(* IEC 61131-3 sources: 2026_Projet_YGO_ExcavatriceDragage/TOOLS/TEST_AUTO_CI/RESULTS/L_SIMULATION/tests (part 7) *)

TEST 'TC-T418-INT-002 Refus puis retour permis sans nouvel appui'
nx := 5000; ny := 5000; raw1 := 0; raw2 := 0; previousButton := FALSE; buttonEdges := 0;
bench.Enable := TRUE; joy.Enable := TRUE; joy.ArmingPermit := TRUE; diagOk.Operational := TRUE;
joy.BusCanOpenOP := diagOk; joy.JoystickOP := diagOk; home.Enable := TRUE; home.BootReady := TRUE;
home.Mode := E_Mode.MAINT_N1; home.BucketOffsetValid := TRUE; home.WinchesMechanicallyStopped := TRUE;
joy.ArmingPermit := FALSE;
ADVANCE_TIME(10000000);
bench(RawPosM1 := raw1, RawPosM2 := raw2);
joy(RawX := bench.Operator.JoyXRaw_ANA1, RawY := bench.Operator.JoyYRaw_ANA2, RawButton := bench.Operator.JoyBtnRaw, Cfg := cfg, NeutralXMem := nx, NeutralYMem := ny);
home(DeadmanArmed := joy.DeadmanArmed, JoystickDeflected := NOT joy.AtNeutralXY, JoystickPull := joy.AxisCmdY.DirectionPositive, JoystickPush := joy.AxisCmdY.DirectionNegative, BtnValidation := bench.Operator.JoyBtnRaw);
IF bench.Operator.JoyBtnRaw AND NOT previousButton THEN buttonEdges := buttonEdges + 1; END_IF; previousButton := bench.Operator.JoyBtnRaw;
bench.SimJoystickFwd_Up_Close_Active := TRUE;
ADVANCE_TIME(10000000);
bench(RawPosM1 := raw1, RawPosM2 := raw2);
joy(RawX := bench.Operator.JoyXRaw_ANA1, RawY := bench.Operator.JoyYRaw_ANA2, RawButton := bench.Operator.JoyBtnRaw, Cfg := cfg, NeutralXMem := nx, NeutralYMem := ny);
home(DeadmanArmed := joy.DeadmanArmed, JoystickDeflected := NOT joy.AtNeutralXY, JoystickPull := joy.AxisCmdY.DirectionPositive, JoystickPush := joy.AxisCmdY.DirectionNegative, BtnValidation := bench.Operator.JoyBtnRaw);
IF bench.Operator.JoyBtnRaw AND NOT previousButton THEN buttonEdges := buttonEdges + 1; END_IF; previousButton := bench.Operator.JoyBtnRaw;
ASSERT_FALSE(joy.AxisCmdY.StartStop, 'Permis absent aucun mouvement'); ASSERT_FALSE(joy.DeadmanArmed, 'Refus reel');
ADVANCE_TIME(10000000);
bench(RawPosM1 := raw1, RawPosM2 := raw2);
joy(RawX := bench.Operator.JoyXRaw_ANA1, RawY := bench.Operator.JoyYRaw_ANA2, RawButton := bench.Operator.JoyBtnRaw, Cfg := cfg, NeutralXMem := nx, NeutralYMem := ny);
home(DeadmanArmed := joy.DeadmanArmed, JoystickDeflected := NOT joy.AtNeutralXY, JoystickPull := joy.AxisCmdY.DirectionPositive, JoystickPush := joy.AxisCmdY.DirectionNegative, BtnValidation := bench.Operator.JoyBtnRaw);
IF bench.Operator.JoyBtnRaw AND NOT previousButton THEN buttonEdges := buttonEdges + 1; END_IF; previousButton := bench.Operator.JoyBtnRaw;
ASSERT_FALSE(joy.AxisCmdY.StartStop, 'Permis absent aucun mouvement'); ASSERT_FALSE(joy.DeadmanArmed, 'Refus reel');
ADVANCE_TIME(10000000);
bench(RawPosM1 := raw1, RawPosM2 := raw2);
joy(RawX := bench.Operator.JoyXRaw_ANA1, RawY := bench.Operator.JoyYRaw_ANA2, RawButton := bench.Operator.JoyBtnRaw, Cfg := cfg, NeutralXMem := nx, NeutralYMem := ny);
home(DeadmanArmed := joy.DeadmanArmed, JoystickDeflected := NOT joy.AtNeutralXY, JoystickPull := joy.AxisCmdY.DirectionPositive, JoystickPush := joy.AxisCmdY.DirectionNegative, BtnValidation := bench.Operator.JoyBtnRaw);
IF bench.Operator.JoyBtnRaw AND NOT previousButton THEN buttonEdges := buttonEdges + 1; END_IF; previousButton := bench.Operator.JoyBtnRaw;
ASSERT_FALSE(joy.AxisCmdY.StartStop, 'Permis absent aucun mouvement'); ASSERT_FALSE(joy.DeadmanArmed, 'Refus reel');
ADVANCE_TIME(10000000);
bench(RawPosM1 := raw1, RawPosM2 := raw2);
joy(RawX := bench.Operator.JoyXRaw_ANA1, RawY := bench.Operator.JoyYRaw_ANA2, RawButton := bench.Operator.JoyBtnRaw, Cfg := cfg, NeutralXMem := nx, NeutralYMem := ny);
home(DeadmanArmed := joy.DeadmanArmed, JoystickDeflected := NOT joy.AtNeutralXY, JoystickPull := joy.AxisCmdY.DirectionPositive, JoystickPush := joy.AxisCmdY.DirectionNegative, BtnValidation := bench.Operator.JoyBtnRaw);
IF bench.Operator.JoyBtnRaw AND NOT previousButton THEN buttonEdges := buttonEdges + 1; END_IF; previousButton := bench.Operator.JoyBtnRaw;
ASSERT_FALSE(joy.AxisCmdY.StartStop, 'Permis absent aucun mouvement'); ASSERT_FALSE(joy.DeadmanArmed, 'Refus reel');
ADVANCE_TIME(10000000);
bench(RawPosM1 := raw1, RawPosM2 := raw2);
joy(RawX := bench.Operator.JoyXRaw_ANA1, RawY := bench.Operator.JoyYRaw_ANA2, RawButton := bench.Operator.JoyBtnRaw, Cfg := cfg, NeutralXMem := nx, NeutralYMem := ny);
home(DeadmanArmed := joy.DeadmanArmed, JoystickDeflected := NOT joy.AtNeutralXY, JoystickPull := joy.AxisCmdY.DirectionPositive, JoystickPush := joy.AxisCmdY.DirectionNegative, BtnValidation := bench.Operator.JoyBtnRaw);
IF bench.Operator.JoyBtnRaw AND NOT previousButton THEN buttonEdges := buttonEdges + 1; END_IF; previousButton := bench.Operator.JoyBtnRaw;
ASSERT_FALSE(joy.AxisCmdY.StartStop, 'Permis absent aucun mouvement'); ASSERT_FALSE(joy.DeadmanArmed, 'Refus reel');
ADVANCE_TIME(10000000);
bench(RawPosM1 := raw1, RawPosM2 := raw2);
joy(RawX := bench.Operator.JoyXRaw_ANA1, RawY := bench.Operator.JoyYRaw_ANA2, RawButton := bench.Operator.JoyBtnRaw, Cfg := cfg, NeutralXMem := nx, NeutralYMem := ny);
home(DeadmanArmed := joy.DeadmanArmed, JoystickDeflected := NOT joy.AtNeutralXY, JoystickPull := joy.AxisCmdY.DirectionPositive, JoystickPush := joy.AxisCmdY.DirectionNegative, BtnValidation := bench.Operator.JoyBtnRaw);
IF bench.Operator.JoyBtnRaw AND NOT previousButton THEN buttonEdges := buttonEdges + 1; END_IF; previousButton := bench.Operator.JoyBtnRaw;
ASSERT_FALSE(joy.AxisCmdY.StartStop, 'Permis absent aucun mouvement'); ASSERT_FALSE(joy.DeadmanArmed, 'Refus reel');
ADVANCE_TIME(10000000);
bench(RawPosM1 := raw1, RawPosM2 := raw2);
joy(RawX := bench.Operator.JoyXRaw_ANA1, RawY := bench.Operator.JoyYRaw_ANA2, RawButton := bench.Operator.JoyBtnRaw, Cfg := cfg, NeutralXMem := nx, NeutralYMem := ny);
home(DeadmanArmed := joy.DeadmanArmed, JoystickDeflected := NOT joy.AtNeutralXY, JoystickPull := joy.AxisCmdY.DirectionPositive, JoystickPush := joy.AxisCmdY.DirectionNegative, BtnValidation := bench.Operator.JoyBtnRaw);
IF bench.Operator.JoyBtnRaw AND NOT previousButton THEN buttonEdges := buttonEdges + 1; END_IF; previousButton := bench.Operator.JoyBtnRaw;
ASSERT_FALSE(joy.AxisCmdY.StartStop, 'Permis absent aucun mouvement'); ASSERT_FALSE(joy.DeadmanArmed, 'Refus reel');
ADVANCE_TIME(10000000);
bench(RawPosM1 := raw1, RawPosM2 := raw2);
joy(RawX := bench.Operator.JoyXRaw_ANA1, RawY := bench.Operator.JoyYRaw_ANA2, RawButton := bench.Operator.JoyBtnRaw, Cfg := cfg, NeutralXMem := nx, NeutralYMem := ny);
home(DeadmanArmed := joy.DeadmanArmed, JoystickDeflected := NOT joy.AtNeutralXY, JoystickPull := joy.AxisCmdY.DirectionPositive, JoystickPush := joy.AxisCmdY.DirectionNegative, BtnValidation := bench.Operator.JoyBtnRaw);
IF bench.Operator.JoyBtnRaw AND NOT previousButton THEN buttonEdges := buttonEdges + 1; END_IF; previousButton := bench.Operator.JoyBtnRaw;
ASSERT_FALSE(joy.AxisCmdY.StartStop, 'Permis absent aucun mouvement'); ASSERT_FALSE(joy.DeadmanArmed, 'Refus reel');
ADVANCE_TIME(10000000);
bench(RawPosM1 := raw1, RawPosM2 := raw2);
joy(RawX := bench.Operator.JoyXRaw_ANA1, RawY := bench.Operator.JoyYRaw_ANA2, RawButton := bench.Operator.JoyBtnRaw, Cfg := cfg, NeutralXMem := nx, NeutralYMem := ny);
home(DeadmanArmed := joy.DeadmanArmed, JoystickDeflected := NOT joy.AtNeutralXY, JoystickPull := joy.AxisCmdY.DirectionPositive, JoystickPush := joy.AxisCmdY.DirectionNegative, BtnValidation := bench.Operator.JoyBtnRaw);
IF bench.Operator.JoyBtnRaw AND NOT previousButton THEN buttonEdges := buttonEdges + 1; END_IF; previousButton := bench.Operator.JoyBtnRaw;
ASSERT_FALSE(joy.AxisCmdY.StartStop, 'Permis absent aucun mouvement'); ASSERT_FALSE(joy.DeadmanArmed, 'Refus reel');
ADVANCE_TIME(10000000);
bench(RawPosM1 := raw1, RawPosM2 := raw2);
joy(RawX := bench.Operator.JoyXRaw_ANA1, RawY := bench.Operator.JoyYRaw_ANA2, RawButton := bench.Operator.JoyBtnRaw, Cfg := cfg, NeutralXMem := nx, NeutralYMem := ny);
home(DeadmanArmed := joy.DeadmanArmed, JoystickDeflected := NOT joy.AtNeutralXY, JoystickPull := joy.AxisCmdY.DirectionPositive, JoystickPush := joy.AxisCmdY.DirectionNegative, BtnValidation := bench.Operator.JoyBtnRaw);
IF bench.Operator.JoyBtnRaw AND NOT previousButton THEN buttonEdges := buttonEdges + 1; END_IF; previousButton := bench.Operator.JoyBtnRaw;
ASSERT_FALSE(joy.AxisCmdY.StartStop, 'Permis absent aucun mouvement'); ASSERT_FALSE(joy.DeadmanArmed, 'Refus reel');
ADVANCE_TIME(10000000);
bench(RawPosM1 := raw1, RawPosM2 := raw2);
joy(RawX := bench.Operator.JoyXRaw_ANA1, RawY := bench.Operator.JoyYRaw_ANA2, RawButton := bench.Operator.JoyBtnRaw, Cfg := cfg, NeutralXMem := nx, NeutralYMem := ny);
home(DeadmanArmed := joy.DeadmanArmed, JoystickDeflected := NOT joy.AtNeutralXY, JoystickPull := joy.AxisCmdY.DirectionPositive, JoystickPush := joy.AxisCmdY.DirectionNegative, BtnValidation := bench.Operator.JoyBtnRaw);
IF bench.Operator.JoyBtnRaw AND NOT previousButton THEN buttonEdges := buttonEdges + 1; END_IF; previousButton := bench.Operator.JoyBtnRaw;
ASSERT_FALSE(joy.AxisCmdY.StartStop, 'Permis absent aucun mouvement'); ASSERT_FALSE(joy.DeadmanArmed, 'Refus reel');
ADVANCE_TIME(10000000);
bench(RawPosM1 := raw1, RawPosM2 := raw2);
joy(RawX := bench.Operator.JoyXRaw_ANA1, RawY := bench.Operator.JoyYRaw_ANA2, RawButton := bench.Operator.JoyBtnRaw, Cfg := cfg, NeutralXMem := nx, NeutralYMem := ny);
home(DeadmanArmed := joy.DeadmanArmed, JoystickDeflected := NOT joy.AtNeutralXY, JoystickPull := joy.AxisCmdY.DirectionPositive, JoystickPush := joy.AxisCmdY.DirectionNegative, BtnValidation := bench.Operator.JoyBtnRaw);
IF bench.Operator.JoyBtnRaw AND NOT previousButton THEN buttonEdges := buttonEdges + 1; END_IF; previousButton := bench.Operator.JoyBtnRaw;
ASSERT_FALSE(joy.AxisCmdY.StartStop, 'Permis absent aucun mouvement'); ASSERT_FALSE(joy.DeadmanArmed, 'Refus reel');
ADVANCE_TIME(10000000);
bench(RawPosM1 := raw1, RawPosM2 := raw2);
joy(RawX := bench.Operator.JoyXRaw_ANA1, RawY := bench.Operator.JoyYRaw_ANA2, RawButton := bench.Operator.JoyBtnRaw, Cfg := cfg, NeutralXMem := nx, NeutralYMem := ny);
home(DeadmanArmed := joy.DeadmanArmed, JoystickDeflected := NOT joy.AtNeutralXY, JoystickPull := joy.AxisCmdY.DirectionPositive, JoystickPush := joy.AxisCmdY.DirectionNegative, BtnValidation := bench.Operator.JoyBtnRaw);
IF bench.Operator.JoyBtnRaw AND NOT previousButton THEN buttonEdges := buttonEdges + 1; END_IF; previousButton := bench.Operator.JoyBtnRaw;
ASSERT_FALSE(joy.AxisCmdY.StartStop, 'Permis absent aucun mouvement'); ASSERT_FALSE(joy.DeadmanArmed, 'Refus reel');
ADVANCE_TIME(10000000);
bench(RawPosM1 := raw1, RawPosM2 := raw2);
joy(RawX := bench.Operator.JoyXRaw_ANA1, RawY := bench.Operator.JoyYRaw_ANA2, RawButton := bench.Operator.JoyBtnRaw, Cfg := cfg, NeutralXMem := nx, NeutralYMem := ny);
home(DeadmanArmed := joy.DeadmanArmed, JoystickDeflected := NOT joy.AtNeutralXY, JoystickPull := joy.AxisCmdY.DirectionPositive, JoystickPush := joy.AxisCmdY.DirectionNegative, BtnValidation := bench.Operator.JoyBtnRaw);
IF bench.Operator.JoyBtnRaw AND NOT previousButton THEN buttonEdges := buttonEdges + 1; END_IF; previousButton := bench.Operator.JoyBtnRaw;
ASSERT_FALSE(joy.AxisCmdY.StartStop, 'Permis absent aucun mouvement'); ASSERT_FALSE(joy.DeadmanArmed, 'Refus reel');
ADVANCE_TIME(10000000);
bench(RawPosM1 := raw1, RawPosM2 := raw2);
joy(RawX := bench.Operator.JoyXRaw_ANA1, RawY := bench.Operator.JoyYRaw_ANA2, RawButton := bench.Operator.JoyBtnRaw, Cfg := cfg, NeutralXMem := nx, NeutralYMem := ny);
home(DeadmanArmed := joy.DeadmanArmed, JoystickDeflected := NOT joy.AtNeutralXY, JoystickPull := joy.AxisCmdY.DirectionPositive, JoystickPush := joy.AxisCmdY.DirectionNegative, BtnValidation := bench.Operator.JoyBtnRaw);
IF bench.Operator.JoyBtnRaw AND NOT previousButton THEN buttonEdges := buttonEdges + 1; END_IF; previousButton := bench.Operator.JoyBtnRaw;
ASSERT_FALSE(joy.AxisCmdY.StartStop, 'Permis absent aucun mouvement'); ASSERT_FALSE(joy.DeadmanArmed, 'Refus reel');
ADVANCE_TIME(10000000);
bench(RawPosM1 := raw1, RawPosM2 := raw2);
joy(RawX := bench.Operator.JoyXRaw_ANA1, RawY := bench.Operator.JoyYRaw_ANA2, RawButton := bench.Operator.JoyBtnRaw, Cfg := cfg, NeutralXMem := nx, NeutralYMem := ny);
home(DeadmanArmed := joy.DeadmanArmed, JoystickDeflected := NOT joy.AtNeutralXY, JoystickPull := joy.AxisCmdY.DirectionPositive, JoystickPush := joy.AxisCmdY.DirectionNegative, BtnValidation := bench.Operator.JoyBtnRaw);
IF bench.Operator.JoyBtnRaw AND NOT previousButton THEN buttonEdges := buttonEdges + 1; END_IF; previousButton := bench.Operator.JoyBtnRaw;
ASSERT_FALSE(joy.AxisCmdY.StartStop, 'Permis absent aucun mouvement'); ASSERT_FALSE(joy.DeadmanArmed, 'Refus reel');
ADVANCE_TIME(10000000);
bench(RawPosM1 := raw1, RawPosM2 := raw2);
joy(RawX := bench.Operator.JoyXRaw_ANA1, RawY := bench.Operator.JoyYRaw_ANA2, RawButton := bench.Operator.JoyBtnRaw, Cfg := cfg, NeutralXMem := nx, NeutralYMem := ny);
home(DeadmanArmed := joy.DeadmanArmed, JoystickDeflected := NOT joy.AtNeutralXY, JoystickPull := joy.AxisCmdY.DirectionPositive, JoystickPush := joy.AxisCmdY.DirectionNegative, BtnValidation := bench.Operator.JoyBtnRaw);
IF bench.Operator.JoyBtnRaw AND NOT previousButton THEN buttonEdges := buttonEdges + 1; END_IF; previousButton := bench.Operator.JoyBtnRaw;
ASSERT_FALSE(joy.AxisCmdY.StartStop, 'Permis absent aucun mouvement'); ASSERT_FALSE(joy.DeadmanArmed, 'Refus reel');
ADVANCE_TIME(10000000);
bench(RawPosM1 := raw1, RawPosM2 := raw2);
joy(RawX := bench.Operator.JoyXRaw_ANA1, RawY := bench.Operator.JoyYRaw_ANA2, RawButton := bench.Operator.JoyBtnRaw, Cfg := cfg, NeutralXMem := nx, NeutralYMem := ny);
home(DeadmanArmed := joy.DeadmanArmed, JoystickDeflected := NOT joy.AtNeutralXY, JoystickPull := joy.AxisCmdY.DirectionPositive, JoystickPush := joy.AxisCmdY.DirectionNegative, BtnValidation := bench.Operator.JoyBtnRaw);
IF bench.Operator.JoyBtnRaw AND NOT previousButton THEN buttonEdges := buttonEdges + 1; END_IF; previousButton := bench.Operator.JoyBtnRaw;
ASSERT_FALSE(joy.AxisCmdY.StartStop, 'Permis absent aucun mouvement'); ASSERT_FALSE(joy.DeadmanArmed, 'Refus reel');
ADVANCE_TIME(10000000);
bench(RawPosM1 := raw1, RawPosM2 := raw2);
joy(RawX := bench.Operator.JoyXRaw_ANA1, RawY := bench.Operator.JoyYRaw_ANA2, RawButton := bench.Operator.JoyBtnRaw, Cfg := cfg, NeutralXMem := nx, NeutralYMem := ny);
home(DeadmanArmed := joy.DeadmanArmed, JoystickDeflected := NOT joy.AtNeutralXY, JoystickPull := joy.AxisCmdY.DirectionPositive, JoystickPush := joy.AxisCmdY.DirectionNegative, BtnValidation := bench.Operator.JoyBtnRaw);
IF bench.Operator.JoyBtnRaw AND NOT previousButton THEN buttonEdges := buttonEdges + 1; END_IF; previousButton := bench.Operator.JoyBtnRaw;
ASSERT_FALSE(joy.AxisCmdY.StartStop, 'Permis absent aucun mouvement'); ASSERT_FALSE(joy.DeadmanArmed, 'Refus reel');
ADVANCE_TIME(10000000);
bench(RawPosM1 := raw1, RawPosM2 := raw2);
joy(RawX := bench.Operator.JoyXRaw_ANA1, RawY := bench.Operator.JoyYRaw_ANA2, RawButton := bench.Operator.JoyBtnRaw, Cfg := cfg, NeutralXMem := nx, NeutralYMem := ny);
home(DeadmanArmed := joy.DeadmanArmed, JoystickDeflected := NOT joy.AtNeutralXY, JoystickPull := joy.AxisCmdY.DirectionPositive, JoystickPush := joy.AxisCmdY.DirectionNegative, BtnValidation := bench.Operator.JoyBtnRaw);
IF bench.Operator.JoyBtnRaw AND NOT previousButton THEN buttonEdges := buttonEdges + 1; END_IF; previousButton := bench.Operator.JoyBtnRaw;
ASSERT_FALSE(joy.AxisCmdY.StartStop, 'Permis absent aucun mouvement'); ASSERT_FALSE(joy.DeadmanArmed, 'Refus reel');
ADVANCE_TIME(10000000);
bench(RawPosM1 := raw1, RawPosM2 := raw2);
joy(RawX := bench.Operator.JoyXRaw_ANA1, RawY := bench.Operator.JoyYRaw_ANA2, RawButton := bench.Operator.JoyBtnRaw, Cfg := cfg, NeutralXMem := nx, NeutralYMem := ny);
home(DeadmanArmed := joy.DeadmanArmed, JoystickDeflected := NOT joy.AtNeutralXY, JoystickPull := joy.AxisCmdY.DirectionPositive, JoystickPush := joy.AxisCmdY.DirectionNegative, BtnValidation := bench.Operator.JoyBtnRaw);
IF bench.Operator.JoyBtnRaw AND NOT previousButton THEN buttonEdges := buttonEdges + 1; END_IF; previousButton := bench.Operator.JoyBtnRaw;
ASSERT_FALSE(joy.AxisCmdY.StartStop, 'Permis absent aucun mouvement'); ASSERT_FALSE(joy.DeadmanArmed, 'Refus reel');
ADVANCE_TIME(10000000);
bench(RawPosM1 := raw1, RawPosM2 := raw2);
joy(RawX := bench.Operator.JoyXRaw_ANA1, RawY := bench.Operator.JoyYRaw_ANA2, RawButton := bench.Operator.JoyBtnRaw, Cfg := cfg, NeutralXMem := nx, NeutralYMem := ny);
home(DeadmanArmed := joy.DeadmanArmed, JoystickDeflected := NOT joy.AtNeutralXY, JoystickPull := joy.AxisCmdY.DirectionPositive, JoystickPush := joy.AxisCmdY.DirectionNegative, BtnValidation := bench.Operator.JoyBtnRaw);
IF bench.Operator.JoyBtnRaw AND NOT previousButton THEN buttonEdges := buttonEdges + 1; END_IF; previousButton := bench.Operator.JoyBtnRaw;
ASSERT_FALSE(joy.AxisCmdY.StartStop, 'Permis absent aucun mouvement'); ASSERT_FALSE(joy.DeadmanArmed, 'Refus reel');
ADVANCE_TIME(10000000);
bench(RawPosM1 := raw1, RawPosM2 := raw2);
joy(RawX := bench.Operator.JoyXRaw_ANA1, RawY := bench.Operator.JoyYRaw_ANA2, RawButton := bench.Operator.JoyBtnRaw, Cfg := cfg, NeutralXMem := nx, NeutralYMem := ny);
home(DeadmanArmed := joy.DeadmanArmed, JoystickDeflected := NOT joy.AtNeutralXY, JoystickPull := joy.AxisCmdY.DirectionPositive, JoystickPush := joy.AxisCmdY.DirectionNegative, BtnValidation := bench.Operator.JoyBtnRaw);
IF bench.Operator.JoyBtnRaw AND NOT previousButton THEN buttonEdges := buttonEdges + 1; END_IF; previousButton := bench.Operator.JoyBtnRaw;
ASSERT_FALSE(joy.AxisCmdY.StartStop, 'Permis absent aucun mouvement'); ASSERT_FALSE(joy.DeadmanArmed, 'Refus reel');
ADVANCE_TIME(10000000);
bench(RawPosM1 := raw1, RawPosM2 := raw2);
joy(RawX := bench.Operator.JoyXRaw_ANA1, RawY := bench.Operator.JoyYRaw_ANA2, RawButton := bench.Operator.JoyBtnRaw, Cfg := cfg, NeutralXMem := nx, NeutralYMem := ny);
home(DeadmanArmed := joy.DeadmanArmed, JoystickDeflected := NOT joy.AtNeutralXY, JoystickPull := joy.AxisCmdY.DirectionPositive, JoystickPush := joy.AxisCmdY.DirectionNegative, BtnValidation := bench.Operator.JoyBtnRaw);
IF bench.Operator.JoyBtnRaw AND NOT previousButton THEN buttonEdges := buttonEdges + 1; END_IF; previousButton := bench.Operator.JoyBtnRaw;
ASSERT_FALSE(joy.AxisCmdY.StartStop, 'Permis absent aucun mouvement'); ASSERT_FALSE(joy.DeadmanArmed, 'Refus reel');
ADVANCE_TIME(10000000);
bench(RawPosM1 := raw1, RawPosM2 := raw2);
joy(RawX := bench.Operator.JoyXRaw_ANA1, RawY := bench.Operator.JoyYRaw_ANA2, RawButton := bench.Operator.JoyBtnRaw, Cfg := cfg, NeutralXMem := nx, NeutralYMem := ny);
home(DeadmanArmed := joy.DeadmanArmed, JoystickDeflected := NOT joy.AtNeutralXY, JoystickPull := joy.AxisCmdY.DirectionPositive, JoystickPush := joy.AxisCmdY.DirectionNegative, BtnValidation := bench.Operator.JoyBtnRaw);
IF bench.Operator.JoyBtnRaw AND NOT previousButton THEN buttonEdges := buttonEdges + 1; END_IF; previousButton := bench.Operator.JoyBtnRaw;
ASSERT_FALSE(joy.AxisCmdY.StartStop, 'Permis absent aucun mouvement'); ASSERT_FALSE(joy.DeadmanArmed, 'Refus reel');
ADVANCE_TIME(10000000);
bench(RawPosM1 := raw1, RawPosM2 := raw2);
joy(RawX := bench.Operator.JoyXRaw_ANA1, RawY := bench.Operator.JoyYRaw_ANA2, RawButton := bench.Operator.JoyBtnRaw, Cfg := cfg, NeutralXMem := nx, NeutralYMem := ny);
home(DeadmanArmed := joy.DeadmanArmed, JoystickDeflected := NOT joy.AtNeutralXY, JoystickPull := joy.AxisCmdY.DirectionPositive, JoystickPush := joy.AxisCmdY.DirectionNegative, BtnValidation := bench.Operator.JoyBtnRaw);
IF bench.Operator.JoyBtnRaw AND NOT previousButton THEN buttonEdges := buttonEdges + 1; END_IF; previousButton := bench.Operator.JoyBtnRaw;
ASSERT_FALSE(joy.AxisCmdY.StartStop, 'Permis absent aucun mouvement'); ASSERT_FALSE(joy.DeadmanArmed, 'Refus reel');
ADVANCE_TIME(10000000);
bench(RawPosM1 := raw1, RawPosM2 := raw2);
joy(RawX := bench.Operator.JoyXRaw_ANA1, RawY := bench.Operator.JoyYRaw_ANA2, RawButton := bench.Operator.JoyBtnRaw, Cfg := cfg, NeutralXMem := nx, NeutralYMem := ny);
home(DeadmanArmed := joy.DeadmanArmed, JoystickDeflected := NOT joy.AtNeutralXY, JoystickPull := joy.AxisCmdY.DirectionPositive, JoystickPush := joy.AxisCmdY.DirectionNegative, BtnValidation := bench.Operator.JoyBtnRaw);
IF bench.Operator.JoyBtnRaw AND NOT previousButton THEN buttonEdges := buttonEdges + 1; END_IF; previousButton := bench.Operator.JoyBtnRaw;
ASSERT_FALSE(joy.AxisCmdY.StartStop, 'Permis absent aucun mouvement'); ASSERT_FALSE(joy.DeadmanArmed, 'Refus reel');
ADVANCE_TIME(10000000);
bench(RawPosM1 := raw1, RawPosM2 := raw2);
joy(RawX := bench.Operator.JoyXRaw_ANA1, RawY := bench.Operator.JoyYRaw_ANA2, RawButton := bench.Operator.JoyBtnRaw, Cfg := cfg, NeutralXMem := nx, NeutralYMem := ny);
home(DeadmanArmed := joy.DeadmanArmed, JoystickDeflected := NOT joy.AtNeutralXY, JoystickPull := joy.AxisCmdY.DirectionPositive, JoystickPush := joy.AxisCmdY.DirectionNegative, BtnValidation := bench.Operator.JoyBtnRaw);
IF bench.Operator.JoyBtnRaw AND NOT previousButton THEN buttonEdges := buttonEdges + 1; END_IF; previousButton := bench.Operator.JoyBtnRaw;
ASSERT_FALSE(joy.AxisCmdY.StartStop, 'Permis absent aucun mouvement'); ASSERT_FALSE(joy.DeadmanArmed, 'Refus reel');
ADVANCE_TIME(10000000);
bench(RawPosM1 := raw1, RawPosM2 := raw2);
joy(RawX := bench.Operator.JoyXRaw_ANA1, RawY := bench.Operator.JoyYRaw_ANA2, RawButton := bench.Operator.JoyBtnRaw, Cfg := cfg, NeutralXMem := nx, NeutralYMem := ny);
home(DeadmanArmed := joy.DeadmanArmed, JoystickDeflected := NOT joy.AtNeutralXY, JoystickPull := joy.AxisCmdY.DirectionPositive, JoystickPush := joy.AxisCmdY.DirectionNegative, BtnValidation := bench.Operator.JoyBtnRaw);
IF bench.Operator.JoyBtnRaw AND NOT previousButton THEN buttonEdges := buttonEdges + 1; END_IF; previousButton := bench.Operator.JoyBtnRaw;
ASSERT_FALSE(joy.AxisCmdY.StartStop, 'Permis absent aucun mouvement'); ASSERT_FALSE(joy.DeadmanArmed, 'Refus reel');
ADVANCE_TIME(10000000);
bench(RawPosM1 := raw1, RawPosM2 := raw2);
joy(RawX := bench.Operator.JoyXRaw_ANA1, RawY := bench.Operator.JoyYRaw_ANA2, RawButton := bench.Operator.JoyBtnRaw, Cfg := cfg, NeutralXMem := nx, NeutralYMem := ny);
home(DeadmanArmed := joy.DeadmanArmed, JoystickDeflected := NOT joy.AtNeutralXY, JoystickPull := joy.AxisCmdY.DirectionPositive, JoystickPush := joy.AxisCmdY.DirectionNegative, BtnValidation := bench.Operator.JoyBtnRaw);
IF bench.Operator.JoyBtnRaw AND NOT previousButton THEN buttonEdges := buttonEdges + 1; END_IF; previousButton := bench.Operator.JoyBtnRaw;
ASSERT_FALSE(joy.AxisCmdY.StartStop, 'Permis absent aucun mouvement'); ASSERT_FALSE(joy.DeadmanArmed, 'Refus reel');
ADVANCE_TIME(10000000);
bench(RawPosM1 := raw1, RawPosM2 := raw2);
joy(RawX := bench.Operator.JoyXRaw_ANA1, RawY := bench.Operator.JoyYRaw_ANA2, RawButton := bench.Operator.JoyBtnRaw, Cfg := cfg, NeutralXMem := nx, NeutralYMem := ny);
home(DeadmanArmed := joy.DeadmanArmed, JoystickDeflected := NOT joy.AtNeutralXY, JoystickPull := joy.AxisCmdY.DirectionPositive, JoystickPush := joy.AxisCmdY.DirectionNegative, BtnValidation := bench.Operator.JoyBtnRaw);
IF bench.Operator.JoyBtnRaw AND NOT previousButton THEN buttonEdges := buttonEdges + 1; END_IF; previousButton := bench.Operator.JoyBtnRaw;
ASSERT_FALSE(joy.AxisCmdY.StartStop, 'Permis absent aucun mouvement'); ASSERT_FALSE(joy.DeadmanArmed, 'Refus reel');
ADVANCE_TIME(10000000);
bench(RawPosM1 := raw1, RawPosM2 := raw2);
joy(RawX := bench.Operator.JoyXRaw_ANA1, RawY := bench.Operator.JoyYRaw_ANA2, RawButton := bench.Operator.JoyBtnRaw, Cfg := cfg, NeutralXMem := nx, NeutralYMem := ny);
home(DeadmanArmed := joy.DeadmanArmed, JoystickDeflected := NOT joy.AtNeutralXY, JoystickPull := joy.AxisCmdY.DirectionPositive, JoystickPush := joy.AxisCmdY.DirectionNegative, BtnValidation := bench.Operator.JoyBtnRaw);
IF bench.Operator.JoyBtnRaw AND NOT previousButton THEN buttonEdges := buttonEdges + 1; END_IF; previousButton := bench.Operator.JoyBtnRaw;
ASSERT_FALSE(joy.AxisCmdY.StartStop, 'Permis absent aucun mouvement'); ASSERT_FALSE(joy.DeadmanArmed, 'Refus reel');
ADVANCE_TIME(10000000);
bench(RawPosM1 := raw1, RawPosM2 := raw2);
joy(RawX := bench.Operator.JoyXRaw_ANA1, RawY := bench.Operator.JoyYRaw_ANA2, RawButton := bench.Operator.JoyBtnRaw, Cfg := cfg, NeutralXMem := nx, NeutralYMem := ny);
home(DeadmanArmed := joy.DeadmanArmed, JoystickDeflected := NOT joy.AtNeutralXY, JoystickPull := joy.AxisCmdY.DirectionPositive, JoystickPush := joy.AxisCmdY.DirectionNegative, BtnValidation := bench.Operator.JoyBtnRaw);
IF bench.Operator.JoyBtnRaw AND NOT previousButton THEN buttonEdges := buttonEdges + 1; END_IF; previousButton := bench.Operator.JoyBtnRaw;
ASSERT_FALSE(joy.AxisCmdY.StartStop, 'Permis absent aucun mouvement'); ASSERT_FALSE(joy.DeadmanArmed, 'Refus reel');
ADVANCE_TIME(10000000);
bench(RawPosM1 := raw1, RawPosM2 := raw2);
joy(RawX := bench.Operator.JoyXRaw_ANA1, RawY := bench.Operator.JoyYRaw_ANA2, RawButton := bench.Operator.JoyBtnRaw, Cfg := cfg, NeutralXMem := nx, NeutralYMem := ny);
home(DeadmanArmed := joy.DeadmanArmed, JoystickDeflected := NOT joy.AtNeutralXY, JoystickPull := joy.AxisCmdY.DirectionPositive, JoystickPush := joy.AxisCmdY.DirectionNegative, BtnValidation := bench.Operator.JoyBtnRaw);
IF bench.Operator.JoyBtnRaw AND NOT previousButton THEN buttonEdges := buttonEdges + 1; END_IF; previousButton := bench.Operator.JoyBtnRaw;
ASSERT_FALSE(joy.AxisCmdY.StartStop, 'Permis absent aucun mouvement'); ASSERT_FALSE(joy.DeadmanArmed, 'Refus reel');
ADVANCE_TIME(10000000);
bench(RawPosM1 := raw1, RawPosM2 := raw2);
joy(RawX := bench.Operator.JoyXRaw_ANA1, RawY := bench.Operator.JoyYRaw_ANA2, RawButton := bench.Operator.JoyBtnRaw, Cfg := cfg, NeutralXMem := nx, NeutralYMem := ny);
home(DeadmanArmed := joy.DeadmanArmed, JoystickDeflected := NOT joy.AtNeutralXY, JoystickPull := joy.AxisCmdY.DirectionPositive, JoystickPush := joy.AxisCmdY.DirectionNegative, BtnValidation := bench.Operator.JoyBtnRaw);
IF bench.Operator.JoyBtnRaw AND NOT previousButton THEN buttonEdges := buttonEdges + 1; END_IF; previousButton := bench.Operator.JoyBtnRaw;
ASSERT_FALSE(joy.AxisCmdY.StartStop, 'Permis absent aucun mouvement'); ASSERT_FALSE(joy.DeadmanArmed, 'Refus reel');
ADVANCE_TIME(10000000);
bench(RawPosM1 := raw1, RawPosM2 := raw2);
joy(RawX := bench.Operator.JoyXRaw_ANA1, RawY := bench.Operator.JoyYRaw_ANA2, RawButton := bench.Operator.JoyBtnRaw, Cfg := cfg, NeutralXMem := nx, NeutralYMem := ny);
home(DeadmanArmed := joy.DeadmanArmed, JoystickDeflected := NOT joy.AtNeutralXY, JoystickPull := joy.AxisCmdY.DirectionPositive, JoystickPush := joy.AxisCmdY.DirectionNegative, BtnValidation := bench.Operator.JoyBtnRaw);
IF bench.Operator.JoyBtnRaw AND NOT previousButton THEN buttonEdges := buttonEdges + 1; END_IF; previousButton := bench.Operator.JoyBtnRaw;
ASSERT_FALSE(joy.AxisCmdY.StartStop, 'Permis absent aucun mouvement'); ASSERT_FALSE(joy.DeadmanArmed, 'Refus reel');
ADVANCE_TIME(10000000);
bench(RawPosM1 := raw1, RawPosM2 := raw2);
joy(RawX := bench.Operator.JoyXRaw_ANA1, RawY := bench.Operator.JoyYRaw_ANA2, RawButton := bench.Operator.JoyBtnRaw, Cfg := cfg, NeutralXMem := nx, NeutralYMem := ny);
home(DeadmanArmed := joy.DeadmanArmed, JoystickDeflected := NOT joy.AtNeutralXY, JoystickPull := joy.AxisCmdY.DirectionPositive, JoystickPush := joy.AxisCmdY.DirectionNegative, BtnValidation := bench.Operator.JoyBtnRaw);
IF bench.Operator.JoyBtnRaw AND NOT previousButton THEN buttonEdges := buttonEdges + 1; END_IF; previousButton := bench.Operator.JoyBtnRaw;
ASSERT_FALSE(joy.AxisCmdY.StartStop, 'Permis absent aucun mouvement'); ASSERT_FALSE(joy.DeadmanArmed, 'Refus reel');
ADVANCE_TIME(10000000);
bench(RawPosM1 := raw1, RawPosM2 := raw2);
joy(RawX := bench.Operator.JoyXRaw_ANA1, RawY := bench.Operator.JoyYRaw_ANA2, RawButton := bench.Operator.JoyBtnRaw, Cfg := cfg, NeutralXMem := nx, NeutralYMem := ny);
home(DeadmanArmed := joy.DeadmanArmed, JoystickDeflected := NOT joy.AtNeutralXY, JoystickPull := joy.AxisCmdY.DirectionPositive, JoystickPush := joy.AxisCmdY.DirectionNegative, BtnValidation := bench.Operator.JoyBtnRaw);
IF bench.Operator.JoyBtnRaw AND NOT previousButton THEN buttonEdges := buttonEdges + 1; END_IF; previousButton := bench.Operator.JoyBtnRaw;
ASSERT_FALSE(joy.AxisCmdY.StartStop, 'Permis absent aucun mouvement'); ASSERT_FALSE(joy.DeadmanArmed, 'Refus reel');
ADVANCE_TIME(10000000);
bench(RawPosM1 := raw1, RawPosM2 := raw2);
joy(RawX := bench.Operator.JoyXRaw_ANA1, RawY := bench.Operator.JoyYRaw_ANA2, RawButton := bench.Operator.JoyBtnRaw, Cfg := cfg, NeutralXMem := nx, NeutralYMem := ny);
home(DeadmanArmed := joy.DeadmanArmed, JoystickDeflected := NOT joy.AtNeutralXY, JoystickPull := joy.AxisCmdY.DirectionPositive, JoystickPush := joy.AxisCmdY.DirectionNegative, BtnValidation := bench.Operator.JoyBtnRaw);
IF bench.Operator.JoyBtnRaw AND NOT previousButton THEN buttonEdges := buttonEdges + 1; END_IF; previousButton := bench.Operator.JoyBtnRaw;
ASSERT_FALSE(joy.AxisCmdY.StartStop, 'Permis absent aucun mouvement'); ASSERT_FALSE(joy.DeadmanArmed, 'Refus reel');
ADVANCE_TIME(10000000);
bench(RawPosM1 := raw1, RawPosM2 := raw2);
joy(RawX := bench.Operator.JoyXRaw_ANA1, RawY := bench.Operator.JoyYRaw_ANA2, RawButton := bench.Operator.JoyBtnRaw, Cfg := cfg, NeutralXMem := nx, NeutralYMem := ny);
home(DeadmanArmed := joy.DeadmanArmed, JoystickDeflected := NOT joy.AtNeutralXY, JoystickPull := joy.AxisCmdY.DirectionPositive, JoystickPush := joy.AxisCmdY.DirectionNegative, BtnValidation := bench.Operator.JoyBtnRaw);
IF bench.Operator.JoyBtnRaw AND NOT previousButton THEN buttonEdges := buttonEdges + 1; END_IF; previousButton := bench.Operator.JoyBtnRaw;
ASSERT_FALSE(joy.AxisCmdY.StartStop, 'Permis absent aucun mouvement'); ASSERT_FALSE(joy.DeadmanArmed, 'Refus reel');
ADVANCE_TIME(10000000);
bench(RawPosM1 := raw1, RawPosM2 := raw2);
joy(RawX := bench.Operator.JoyXRaw_ANA1, RawY := bench.Operator.JoyYRaw_ANA2, RawButton := bench.Operator.JoyBtnRaw, Cfg := cfg, NeutralXMem := nx, NeutralYMem := ny);
home(DeadmanArmed := joy.DeadmanArmed, JoystickDeflected := NOT joy.AtNeutralXY, JoystickPull := joy.AxisCmdY.DirectionPositive, JoystickPush := joy.AxisCmdY.DirectionNegative, BtnValidation := bench.Operator.JoyBtnRaw);
IF bench.Operator.JoyBtnRaw AND NOT previousButton THEN buttonEdges := buttonEdges + 1; END_IF; previousButton := bench.Operator.JoyBtnRaw;
ASSERT_FALSE(joy.AxisCmdY.StartStop, 'Permis absent aucun mouvement'); ASSERT_FALSE(joy.DeadmanArmed, 'Refus reel');
ADVANCE_TIME(10000000);
bench(RawPosM1 := raw1, RawPosM2 := raw2);
joy(RawX := bench.Operator.JoyXRaw_ANA1, RawY := bench.Operator.JoyYRaw_ANA2, RawButton := bench.Operator.JoyBtnRaw, Cfg := cfg, NeutralXMem := nx, NeutralYMem := ny);
home(DeadmanArmed := joy.DeadmanArmed, JoystickDeflected := NOT joy.AtNeutralXY, JoystickPull := joy.AxisCmdY.DirectionPositive, JoystickPush := joy.AxisCmdY.DirectionNegative, BtnValidation := bench.Operator.JoyBtnRaw);
IF bench.Operator.JoyBtnRaw AND NOT previousButton THEN buttonEdges := buttonEdges + 1; END_IF; previousButton := bench.Operator.JoyBtnRaw;
ASSERT_FALSE(joy.AxisCmdY.StartStop, 'Permis absent aucun mouvement'); ASSERT_FALSE(joy.DeadmanArmed, 'Refus reel');
ADVANCE_TIME(10000000);
bench(RawPosM1 := raw1, RawPosM2 := raw2);
joy(RawX := bench.Operator.JoyXRaw_ANA1, RawY := bench.Operator.JoyYRaw_ANA2, RawButton := bench.Operator.JoyBtnRaw, Cfg := cfg, NeutralXMem := nx, NeutralYMem := ny);
home(DeadmanArmed := joy.DeadmanArmed, JoystickDeflected := NOT joy.AtNeutralXY, JoystickPull := joy.AxisCmdY.DirectionPositive, JoystickPush := joy.AxisCmdY.DirectionNegative, BtnValidation := bench.Operator.JoyBtnRaw);
IF bench.Operator.JoyBtnRaw AND NOT previousButton THEN buttonEdges := buttonEdges + 1; END_IF; previousButton := bench.Operator.JoyBtnRaw;
ASSERT_FALSE(joy.AxisCmdY.StartStop, 'Permis absent aucun mouvement'); ASSERT_FALSE(joy.DeadmanArmed, 'Refus reel');
ADVANCE_TIME(10000000);
bench(RawPosM1 := raw1, RawPosM2 := raw2);
joy(RawX := bench.Operator.JoyXRaw_ANA1, RawY := bench.Operator.JoyYRaw_ANA2, RawButton := bench.Operator.JoyBtnRaw, Cfg := cfg, NeutralXMem := nx, NeutralYMem := ny);
home(DeadmanArmed := joy.DeadmanArmed, JoystickDeflected := NOT joy.AtNeutralXY, JoystickPull := joy.AxisCmdY.DirectionPositive, JoystickPush := joy.AxisCmdY.DirectionNegative, BtnValidation := bench.Operator.JoyBtnRaw);
IF bench.Operator.JoyBtnRaw AND NOT previousButton THEN buttonEdges := buttonEdges + 1; END_IF; previousButton := bench.Operator.JoyBtnRaw;
ASSERT_FALSE(joy.AxisCmdY.StartStop, 'Permis absent aucun mouvement'); ASSERT_FALSE(joy.DeadmanArmed, 'Refus reel');
ADVANCE_TIME(10000000);
bench(RawPosM1 := raw1, RawPosM2 := raw2);
joy(RawX := bench.Operator.JoyXRaw_ANA1, RawY := bench.Operator.JoyYRaw_ANA2, RawButton := bench.Operator.JoyBtnRaw, Cfg := cfg, NeutralXMem := nx, NeutralYMem := ny);
home(DeadmanArmed := joy.DeadmanArmed, JoystickDeflected := NOT joy.AtNeutralXY, JoystickPull := joy.AxisCmdY.DirectionPositive, JoystickPush := joy.AxisCmdY.DirectionNegative, BtnValidation := bench.Operator.JoyBtnRaw);
IF bench.Operator.JoyBtnRaw AND NOT previousButton THEN buttonEdges := buttonEdges + 1; END_IF; previousButton := bench.Operator.JoyBtnRaw;
ASSERT_FALSE(joy.AxisCmdY.StartStop, 'Permis absent aucun mouvement'); ASSERT_FALSE(joy.DeadmanArmed, 'Refus reel');
ADVANCE_TIME(10000000);
bench(RawPosM1 := raw1, RawPosM2 := raw2);
joy(RawX := bench.Operator.JoyXRaw_ANA1, RawY := bench.Operator.JoyYRaw_ANA2, RawButton := bench.Operator.JoyBtnRaw, Cfg := cfg, NeutralXMem := nx, NeutralYMem := ny);
home(DeadmanArmed := joy.DeadmanArmed, JoystickDeflected := NOT joy.AtNeutralXY, JoystickPull := joy.AxisCmdY.DirectionPositive, JoystickPush := joy.AxisCmdY.DirectionNegative, BtnValidation := bench.Operator.JoyBtnRaw);
IF bench.Operator.JoyBtnRaw AND NOT previousButton THEN buttonEdges := buttonEdges + 1; END_IF; previousButton := bench.Operator.JoyBtnRaw;
ASSERT_FALSE(joy.AxisCmdY.StartStop, 'Permis absent aucun mouvement'); ASSERT_FALSE(joy.DeadmanArmed, 'Refus reel');
ADVANCE_TIME(10000000);
bench(RawPosM1 := raw1, RawPosM2 := raw2);
joy(RawX := bench.Operator.JoyXRaw_ANA1, RawY := bench.Operator.JoyYRaw_ANA2, RawButton := bench.Operator.JoyBtnRaw, Cfg := cfg, NeutralXMem := nx, NeutralYMem := ny);
home(DeadmanArmed := joy.DeadmanArmed, JoystickDeflected := NOT joy.AtNeutralXY, JoystickPull := joy.AxisCmdY.DirectionPositive, JoystickPush := joy.AxisCmdY.DirectionNegative, BtnValidation := bench.Operator.JoyBtnRaw);
IF bench.Operator.JoyBtnRaw AND NOT previousButton THEN buttonEdges := buttonEdges + 1; END_IF; previousButton := bench.Operator.JoyBtnRaw;
ASSERT_FALSE(joy.AxisCmdY.StartStop, 'Permis absent aucun mouvement'); ASSERT_FALSE(joy.DeadmanArmed, 'Refus reel');
ADVANCE_TIME(10000000);
bench(RawPosM1 := raw1, RawPosM2 := raw2);
joy(RawX := bench.Operator.JoyXRaw_ANA1, RawY := bench.Operator.JoyYRaw_ANA2, RawButton := bench.Operator.JoyBtnRaw, Cfg := cfg, NeutralXMem := nx, NeutralYMem := ny);
home(DeadmanArmed := joy.DeadmanArmed, JoystickDeflected := NOT joy.AtNeutralXY, JoystickPull := joy.AxisCmdY.DirectionPositive, JoystickPush := joy.AxisCmdY.DirectionNegative, BtnValidation := bench.Operator.JoyBtnRaw);
IF bench.Operator.JoyBtnRaw AND NOT previousButton THEN buttonEdges := buttonEdges + 1; END_IF; previousButton := bench.Operator.JoyBtnRaw;
ASSERT_FALSE(joy.AxisCmdY.StartStop, 'Permis absent aucun mouvement'); ASSERT_FALSE(joy.DeadmanArmed, 'Refus reel');
ADVANCE_TIME(10000000);
bench(RawPosM1 := raw1, RawPosM2 := raw2);
joy(RawX := bench.Operator.JoyXRaw_ANA1, RawY := bench.Operator.JoyYRaw_ANA2, RawButton := bench.Operator.JoyBtnRaw, Cfg := cfg, NeutralXMem := nx, NeutralYMem := ny);
home(DeadmanArmed := joy.DeadmanArmed, JoystickDeflected := NOT joy.AtNeutralXY, JoystickPull := joy.AxisCmdY.DirectionPositive, JoystickPush := joy.AxisCmdY.DirectionNegative, BtnValidation := bench.Operator.JoyBtnRaw);
IF bench.Operator.JoyBtnRaw AND NOT previousButton THEN buttonEdges := buttonEdges + 1; END_IF; previousButton := bench.Operator.JoyBtnRaw;
ASSERT_FALSE(joy.AxisCmdY.StartStop, 'Permis absent aucun mouvement'); ASSERT_FALSE(joy.DeadmanArmed, 'Refus reel');
ADVANCE_TIME(10000000);
bench(RawPosM1 := raw1, RawPosM2 := raw2);
joy(RawX := bench.Operator.JoyXRaw_ANA1, RawY := bench.Operator.JoyYRaw_ANA2, RawButton := bench.Operator.JoyBtnRaw, Cfg := cfg, NeutralXMem := nx, NeutralYMem := ny);
home(DeadmanArmed := joy.DeadmanArmed, JoystickDeflected := NOT joy.AtNeutralXY, JoystickPull := joy.AxisCmdY.DirectionPositive, JoystickPush := joy.AxisCmdY.DirectionNegative, BtnValidation := bench.Operator.JoyBtnRaw);
IF bench.Operator.JoyBtnRaw AND NOT previousButton THEN buttonEdges := buttonEdges + 1; END_IF; previousButton := bench.Operator.JoyBtnRaw;
ASSERT_FALSE(joy.AxisCmdY.StartStop, 'Permis absent aucun mouvement'); ASSERT_FALSE(joy.DeadmanArmed, 'Refus reel');
ADVANCE_TIME(10000000);
bench(RawPosM1 := raw1, RawPosM2 := raw2);
joy(RawX := bench.Operator.JoyXRaw_ANA1, RawY := bench.Operator.JoyYRaw_ANA2, RawButton := bench.Operator.JoyBtnRaw, Cfg := cfg, NeutralXMem := nx, NeutralYMem := ny);
home(DeadmanArmed := joy.DeadmanArmed, JoystickDeflected := NOT joy.AtNeutralXY, JoystickPull := joy.AxisCmdY.DirectionPositive, JoystickPush := joy.AxisCmdY.DirectionNegative, BtnValidation := bench.Operator.JoyBtnRaw);
IF bench.Operator.JoyBtnRaw AND NOT previousButton THEN buttonEdges := buttonEdges + 1; END_IF; previousButton := bench.Operator.JoyBtnRaw;
ASSERT_FALSE(joy.AxisCmdY.StartStop, 'Permis absent aucun mouvement'); ASSERT_FALSE(joy.DeadmanArmed, 'Refus reel');
ADVANCE_TIME(10000000);
bench(RawPosM1 := raw1, RawPosM2 := raw2);
joy(RawX := bench.Operator.JoyXRaw_ANA1, RawY := bench.Operator.JoyYRaw_ANA2, RawButton := bench.Operator.JoyBtnRaw, Cfg := cfg, NeutralXMem := nx, NeutralYMem := ny);
home(DeadmanArmed := joy.DeadmanArmed, JoystickDeflected := NOT joy.AtNeutralXY, JoystickPull := joy.AxisCmdY.DirectionPositive, JoystickPush := joy.AxisCmdY.DirectionNegative, BtnValidation := bench.Operator.JoyBtnRaw);
IF bench.Operator.JoyBtnRaw AND NOT previousButton THEN buttonEdges := buttonEdges + 1; END_IF; previousButton := bench.Operator.JoyBtnRaw;
ASSERT_FALSE(joy.AxisCmdY.StartStop, 'Permis absent aucun mouvement'); ASSERT_FALSE(joy.DeadmanArmed, 'Refus reel');
ADVANCE_TIME(10000000);
bench(RawPosM1 := raw1, RawPosM2 := raw2);
joy(RawX := bench.Operator.JoyXRaw_ANA1, RawY := bench.Operator.JoyYRaw_ANA2, RawButton := bench.Operator.JoyBtnRaw, Cfg := cfg, NeutralXMem := nx, NeutralYMem := ny);
home(DeadmanArmed := joy.DeadmanArmed, JoystickDeflected := NOT joy.AtNeutralXY, JoystickPull := joy.AxisCmdY.DirectionPositive, JoystickPush := joy.AxisCmdY.DirectionNegative, BtnValidation := bench.Operator.JoyBtnRaw);
IF bench.Operator.JoyBtnRaw AND NOT previousButton THEN buttonEdges := buttonEdges + 1; END_IF; previousButton := bench.Operator.JoyBtnRaw;
ASSERT_FALSE(joy.AxisCmdY.StartStop, 'Permis absent aucun mouvement'); ASSERT_FALSE(joy.DeadmanArmed, 'Refus reel');
ADVANCE_TIME(10000000);
bench(RawPosM1 := raw1, RawPosM2 := raw2);
joy(RawX := bench.Operator.JoyXRaw_ANA1, RawY := bench.Operator.JoyYRaw_ANA2, RawButton := bench.Operator.JoyBtnRaw, Cfg := cfg, NeutralXMem := nx, NeutralYMem := ny);
home(DeadmanArmed := joy.DeadmanArmed, JoystickDeflected := NOT joy.AtNeutralXY, JoystickPull := joy.AxisCmdY.DirectionPositive, JoystickPush := joy.AxisCmdY.DirectionNegative, BtnValidation := bench.Operator.JoyBtnRaw);
IF bench.Operator.JoyBtnRaw AND NOT previousButton THEN buttonEdges := buttonEdges + 1; END_IF; previousButton := bench.Operator.JoyBtnRaw;
ASSERT_FALSE(joy.AxisCmdY.StartStop, 'Permis absent aucun mouvement'); ASSERT_FALSE(joy.DeadmanArmed, 'Refus reel');
ADVANCE_TIME(10000000);
bench(RawPosM1 := raw1, RawPosM2 := raw2);
joy(RawX := bench.Operator.JoyXRaw_ANA1, RawY := bench.Operator.JoyYRaw_ANA2, RawButton := bench.Operator.JoyBtnRaw, Cfg := cfg, NeutralXMem := nx, NeutralYMem := ny);
home(DeadmanArmed := joy.DeadmanArmed, JoystickDeflected := NOT joy.AtNeutralXY, JoystickPull := joy.AxisCmdY.DirectionPositive, JoystickPush := joy.AxisCmdY.DirectionNegative, BtnValidation := bench.Operator.JoyBtnRaw);
IF bench.Operator.JoyBtnRaw AND NOT previousButton THEN buttonEdges := buttonEdges + 1; END_IF; previousButton := bench.Operator.JoyBtnRaw;
ASSERT_FALSE(joy.AxisCmdY.StartStop, 'Permis absent aucun mouvement'); ASSERT_FALSE(joy.DeadmanArmed, 'Refus reel');
ADVANCE_TIME(10000000);
bench(RawPosM1 := raw1, RawPosM2 := raw2);
joy(RawX := bench.Operator.JoyXRaw_ANA1, RawY := bench.Operator.JoyYRaw_ANA2, RawButton := bench.Operator.JoyBtnRaw, Cfg := cfg, NeutralXMem := nx, NeutralYMem := ny);
home(DeadmanArmed := joy.DeadmanArmed, JoystickDeflected := NOT joy.AtNeutralXY, JoystickPull := joy.AxisCmdY.DirectionPositive, JoystickPush := joy.AxisCmdY.DirectionNegative, BtnValidation := bench.Operator.JoyBtnRaw);
IF bench.Operator.JoyBtnRaw AND NOT previousButton THEN buttonEdges := buttonEdges + 1; END_IF; previousButton := bench.Operator.JoyBtnRaw;
ASSERT_FALSE(joy.AxisCmdY.StartStop, 'Permis absent aucun mouvement'); ASSERT_FALSE(joy.DeadmanArmed, 'Refus reel');
ADVANCE_TIME(10000000);
bench(RawPosM1 := raw1, RawPosM2 := raw2);
joy(RawX := bench.Operator.JoyXRaw_ANA1, RawY := bench.Operator.JoyYRaw_ANA2, RawButton := bench.Operator.JoyBtnRaw, Cfg := cfg, NeutralXMem := nx, NeutralYMem := ny);
home(DeadmanArmed := joy.DeadmanArmed, JoystickDeflected := NOT joy.AtNeutralXY, JoystickPull := joy.AxisCmdY.DirectionPositive, JoystickPush := joy.AxisCmdY.DirectionNegative, BtnValidation := bench.Operator.JoyBtnRaw);
IF bench.Operator.JoyBtnRaw AND NOT previousButton THEN buttonEdges := buttonEdges + 1; END_IF; previousButton := bench.Operator.JoyBtnRaw;
ASSERT_FALSE(joy.AxisCmdY.StartStop, 'Permis absent aucun mouvement'); ASSERT_FALSE(joy.DeadmanArmed, 'Refus reel');
ADVANCE_TIME(10000000);
bench(RawPosM1 := raw1, RawPosM2 := raw2);
joy(RawX := bench.Operator.JoyXRaw_ANA1, RawY := bench.Operator.JoyYRaw_ANA2, RawButton := bench.Operator.JoyBtnRaw, Cfg := cfg, NeutralXMem := nx, NeutralYMem := ny);
home(DeadmanArmed := joy.DeadmanArmed, JoystickDeflected := NOT joy.AtNeutralXY, JoystickPull := joy.AxisCmdY.DirectionPositive, JoystickPush := joy.AxisCmdY.DirectionNegative, BtnValidation := bench.Operator.JoyBtnRaw);
IF bench.Operator.JoyBtnRaw AND NOT previousButton THEN buttonEdges := buttonEdges + 1; END_IF; previousButton := bench.Operator.JoyBtnRaw;
ASSERT_FALSE(joy.AxisCmdY.StartStop, 'Permis absent aucun mouvement'); ASSERT_FALSE(joy.DeadmanArmed, 'Refus reel');
ADVANCE_TIME(10000000);
bench(RawPosM1 := raw1, RawPosM2 := raw2);
joy(RawX := bench.Operator.JoyXRaw_ANA1, RawY := bench.Operator.JoyYRaw_ANA2, RawButton := bench.Operator.JoyBtnRaw, Cfg := cfg, NeutralXMem := nx, NeutralYMem := ny);
home(DeadmanArmed := joy.DeadmanArmed, JoystickDeflected := NOT joy.AtNeutralXY, JoystickPull := joy.AxisCmdY.DirectionPositive, JoystickPush := joy.AxisCmdY.DirectionNegative, BtnValidation := bench.Operator.JoyBtnRaw);
IF bench.Operator.JoyBtnRaw AND NOT previousButton THEN buttonEdges := buttonEdges + 1; END_IF; previousButton := bench.Operator.JoyBtnRaw;
ASSERT_FALSE(joy.AxisCmdY.StartStop, 'Permis absent aucun mouvement'); ASSERT_FALSE(joy.DeadmanArmed, 'Refus reel');
ADVANCE_TIME(10000000);
bench(RawPosM1 := raw1, RawPosM2 := raw2);
joy(RawX := bench.Operator.JoyXRaw_ANA1, RawY := bench.Operator.JoyYRaw_ANA2, RawButton := bench.Operator.JoyBtnRaw, Cfg := cfg, NeutralXMem := nx, NeutralYMem := ny);
home(DeadmanArmed := joy.DeadmanArmed, JoystickDeflected := NOT joy.AtNeutralXY, JoystickPull := joy.AxisCmdY.DirectionPositive, JoystickPush := joy.AxisCmdY.DirectionNegative, BtnValidation := bench.Operator.JoyBtnRaw);
IF bench.Operator.JoyBtnRaw AND NOT previousButton THEN buttonEdges := buttonEdges + 1; END_IF; previousButton := bench.Operator.JoyBtnRaw;
ASSERT_FALSE(joy.AxisCmdY.StartStop, 'Permis absent aucun mouvement'); ASSERT_FALSE(joy.DeadmanArmed, 'Refus reel');
ADVANCE_TIME(10000000);
bench(RawPosM1 := raw1, RawPosM2 := raw2);
joy(RawX := bench.Operator.JoyXRaw_ANA1, RawY := bench.Operator.JoyYRaw_ANA2, RawButton := bench.Operator.JoyBtnRaw, Cfg := cfg, NeutralXMem := nx, NeutralYMem := ny);
home(DeadmanArmed := joy.DeadmanArmed, JoystickDeflected := NOT joy.AtNeutralXY, JoystickPull := joy.AxisCmdY.DirectionPositive, JoystickPush := joy.AxisCmdY.DirectionNegative, BtnValidation := bench.Operator.JoyBtnRaw);
IF bench.Operator.JoyBtnRaw AND NOT previousButton THEN buttonEdges := buttonEdges + 1; END_IF; previousButton := bench.Operator.JoyBtnRaw;
ASSERT_FALSE(joy.AxisCmdY.StartStop, 'Permis absent aucun mouvement'); ASSERT_FALSE(joy.DeadmanArmed, 'Refus reel');
ADVANCE_TIME(10000000);
bench(RawPosM1 := raw1, RawPosM2 := raw2);
joy(RawX := bench.Operator.JoyXRaw_ANA1, RawY := bench.Operator.JoyYRaw_ANA2, RawButton := bench.Operator.JoyBtnRaw, Cfg := cfg, NeutralXMem := nx, NeutralYMem := ny);
home(DeadmanArmed := joy.DeadmanArmed, JoystickDeflected := NOT joy.AtNeutralXY, JoystickPull := joy.AxisCmdY.DirectionPositive, JoystickPush := joy.AxisCmdY.DirectionNegative, BtnValidation := bench.Operator.JoyBtnRaw);
IF bench.Operator.JoyBtnRaw AND NOT previousButton THEN buttonEdges := buttonEdges + 1; END_IF; previousButton := bench.Operator.JoyBtnRaw;
ASSERT_FALSE(joy.AxisCmdY.StartStop, 'Permis absent aucun mouvement'); ASSERT_FALSE(joy.DeadmanArmed, 'Refus reel');
ADVANCE_TIME(10000000);
bench(RawPosM1 := raw1, RawPosM2 := raw2);
joy(RawX := bench.Operator.JoyXRaw_ANA1, RawY := bench.Operator.JoyYRaw_ANA2, RawButton := bench.Operator.JoyBtnRaw, Cfg := cfg, NeutralXMem := nx, NeutralYMem := ny);
home(DeadmanArmed := joy.DeadmanArmed, JoystickDeflected := NOT joy.AtNeutralXY, JoystickPull := joy.AxisCmdY.DirectionPositive, JoystickPush := joy.AxisCmdY.DirectionNegative, BtnValidation := bench.Operator.JoyBtnRaw);
IF bench.Operator.JoyBtnRaw AND NOT previousButton THEN buttonEdges := buttonEdges + 1; END_IF; previousButton := bench.Operator.JoyBtnRaw;
ASSERT_FALSE(joy.AxisCmdY.StartStop, 'Permis absent aucun mouvement'); ASSERT_FALSE(joy.DeadmanArmed, 'Refus reel');
ADVANCE_TIME(10000000);
bench(RawPosM1 := raw1, RawPosM2 := raw2);
joy(RawX := bench.Operator.JoyXRaw_ANA1, RawY := bench.Operator.JoyYRaw_ANA2, RawButton := bench.Operator.JoyBtnRaw, Cfg := cfg, NeutralXMem := nx, NeutralYMem := ny);
home(DeadmanArmed := joy.DeadmanArmed, JoystickDeflected := NOT joy.AtNeutralXY, JoystickPull := joy.AxisCmdY.DirectionPositive, JoystickPush := joy.AxisCmdY.DirectionNegative, BtnValidation := bench.Operator.JoyBtnRaw);
IF bench.Operator.JoyBtnRaw AND NOT previousButton THEN buttonEdges := buttonEdges + 1; END_IF; previousButton := bench.Operator.JoyBtnRaw;
ASSERT_FALSE(joy.AxisCmdY.StartStop, 'Permis absent aucun mouvement'); ASSERT_FALSE(joy.DeadmanArmed, 'Refus reel');
ADVANCE_TIME(10000000);
bench(RawPosM1 := raw1, RawPosM2 := raw2);
joy(RawX := bench.Operator.JoyXRaw_ANA1, RawY := bench.Operator.JoyYRaw_ANA2, RawButton := bench.Operator.JoyBtnRaw, Cfg := cfg, NeutralXMem := nx, NeutralYMem := ny);
home(DeadmanArmed := joy.DeadmanArmed, JoystickDeflected := NOT joy.AtNeutralXY, JoystickPull := joy.AxisCmdY.DirectionPositive, JoystickPush := joy.AxisCmdY.DirectionNegative, BtnValidation := bench.Operator.JoyBtnRaw);
IF bench.Operator.JoyBtnRaw AND NOT previousButton THEN buttonEdges := buttonEdges + 1; END_IF; previousButton := bench.Operator.JoyBtnRaw;
ASSERT_FALSE(joy.AxisCmdY.StartStop, 'Permis absent aucun mouvement'); ASSERT_FALSE(joy.DeadmanArmed, 'Refus reel');
joy.ArmingPermit := TRUE;
ADVANCE_TIME(10000000);
bench(RawPosM1 := raw1, RawPosM2 := raw2);
joy(RawX := bench.Operator.JoyXRaw_ANA1, RawY := bench.Operator.JoyYRaw_ANA2, RawButton := bench.Operator.JoyBtnRaw, Cfg := cfg, NeutralXMem := nx, NeutralYMem := ny);
home(DeadmanArmed := joy.DeadmanArmed, JoystickDeflected := NOT joy.AtNeutralXY, JoystickPull := joy.AxisCmdY.DirectionPositive, JoystickPush := joy.AxisCmdY.DirectionNegative, BtnValidation := bench.Operator.JoyBtnRaw);
IF bench.Operator.JoyBtnRaw AND NOT previousButton THEN buttonEdges := buttonEdges + 1; END_IF; previousButton := bench.Operator.JoyBtnRaw;
ASSERT_FALSE(joy.DeadmanArmed, 'Pas de rearmement au retour du permis');
ADVANCE_TIME(10000000);
bench(RawPosM1 := raw1, RawPosM2 := raw2);
joy(RawX := bench.Operator.JoyXRaw_ANA1, RawY := bench.Operator.JoyYRaw_ANA2, RawButton := bench.Operator.JoyBtnRaw, Cfg := cfg, NeutralXMem := nx, NeutralYMem := ny);
home(DeadmanArmed := joy.DeadmanArmed, JoystickDeflected := NOT joy.AtNeutralXY, JoystickPull := joy.AxisCmdY.DirectionPositive, JoystickPush := joy.AxisCmdY.DirectionNegative, BtnValidation := bench.Operator.JoyBtnRaw);
IF bench.Operator.JoyBtnRaw AND NOT previousButton THEN buttonEdges := buttonEdges + 1; END_IF; previousButton := bench.Operator.JoyBtnRaw;
ASSERT_FALSE(joy.DeadmanArmed, 'Pas de rearmement au retour du permis');
ADVANCE_TIME(10000000);
bench(RawPosM1 := raw1, RawPosM2 := raw2);
joy(RawX := bench.Operator.JoyXRaw_ANA1, RawY := bench.Operator.JoyYRaw_ANA2, RawButton := bench.Operator.JoyBtnRaw, Cfg := cfg, NeutralXMem := nx, NeutralYMem := ny);
home(DeadmanArmed := joy.DeadmanArmed, JoystickDeflected := NOT joy.AtNeutralXY, JoystickPull := joy.AxisCmdY.DirectionPositive, JoystickPush := joy.AxisCmdY.DirectionNegative, BtnValidation := bench.Operator.JoyBtnRaw);
IF bench.Operator.JoyBtnRaw AND NOT previousButton THEN buttonEdges := buttonEdges + 1; END_IF; previousButton := bench.Operator.JoyBtnRaw;
ASSERT_FALSE(joy.DeadmanArmed, 'Pas de rearmement au retour du permis');
ADVANCE_TIME(10000000);
bench(RawPosM1 := raw1, RawPosM2 := raw2);
joy(RawX := bench.Operator.JoyXRaw_ANA1, RawY := bench.Operator.JoyYRaw_ANA2, RawButton := bench.Operator.JoyBtnRaw, Cfg := cfg, NeutralXMem := nx, NeutralYMem := ny);
home(DeadmanArmed := joy.DeadmanArmed, JoystickDeflected := NOT joy.AtNeutralXY, JoystickPull := joy.AxisCmdY.DirectionPositive, JoystickPush := joy.AxisCmdY.DirectionNegative, BtnValidation := bench.Operator.JoyBtnRaw);
IF bench.Operator.JoyBtnRaw AND NOT previousButton THEN buttonEdges := buttonEdges + 1; END_IF; previousButton := bench.Operator.JoyBtnRaw;
ASSERT_FALSE(joy.DeadmanArmed, 'Pas de rearmement au retour du permis');
ADVANCE_TIME(10000000);
bench(RawPosM1 := raw1, RawPosM2 := raw2);
joy(RawX := bench.Operator.JoyXRaw_ANA1, RawY := bench.Operator.JoyYRaw_ANA2, RawButton := bench.Operator.JoyBtnRaw, Cfg := cfg, NeutralXMem := nx, NeutralYMem := ny);
home(DeadmanArmed := joy.DeadmanArmed, JoystickDeflected := NOT joy.AtNeutralXY, JoystickPull := joy.AxisCmdY.DirectionPositive, JoystickPush := joy.AxisCmdY.DirectionNegative, BtnValidation := bench.Operator.JoyBtnRaw);
IF bench.Operator.JoyBtnRaw AND NOT previousButton THEN buttonEdges := buttonEdges + 1; END_IF; previousButton := bench.Operator.JoyBtnRaw;
ASSERT_FALSE(joy.DeadmanArmed, 'Pas de rearmement au retour du permis');
ADVANCE_TIME(10000000);
bench(RawPosM1 := raw1, RawPosM2 := raw2);
joy(RawX := bench.Operator.JoyXRaw_ANA1, RawY := bench.Operator.JoyYRaw_ANA2, RawButton := bench.Operator.JoyBtnRaw, Cfg := cfg, NeutralXMem := nx, NeutralYMem := ny);
home(DeadmanArmed := joy.DeadmanArmed, JoystickDeflected := NOT joy.AtNeutralXY, JoystickPull := joy.AxisCmdY.DirectionPositive, JoystickPush := joy.AxisCmdY.DirectionNegative, BtnValidation := bench.Operator.JoyBtnRaw);
IF bench.Operator.JoyBtnRaw AND NOT previousButton THEN buttonEdges := buttonEdges + 1; END_IF; previousButton := bench.Operator.JoyBtnRaw;
ASSERT_FALSE(joy.DeadmanArmed, 'Pas de rearmement au retour du permis');
ADVANCE_TIME(10000000);
bench(RawPosM1 := raw1, RawPosM2 := raw2);
joy(RawX := bench.Operator.JoyXRaw_ANA1, RawY := bench.Operator.JoyYRaw_ANA2, RawButton := bench.Operator.JoyBtnRaw, Cfg := cfg, NeutralXMem := nx, NeutralYMem := ny);
home(DeadmanArmed := joy.DeadmanArmed, JoystickDeflected := NOT joy.AtNeutralXY, JoystickPull := joy.AxisCmdY.DirectionPositive, JoystickPush := joy.AxisCmdY.DirectionNegative, BtnValidation := bench.Operator.JoyBtnRaw);
IF bench.Operator.JoyBtnRaw AND NOT previousButton THEN buttonEdges := buttonEdges + 1; END_IF; previousButton := bench.Operator.JoyBtnRaw;
ASSERT_FALSE(joy.DeadmanArmed, 'Pas de rearmement au retour du permis');
ADVANCE_TIME(10000000);
bench(RawPosM1 := raw1, RawPosM2 := raw2);
joy(RawX := bench.Operator.JoyXRaw_ANA1, RawY := bench.Operator.JoyYRaw_ANA2, RawButton := bench.Operator.JoyBtnRaw, Cfg := cfg, NeutralXMem := nx, NeutralYMem := ny);
home(DeadmanArmed := joy.DeadmanArmed, JoystickDeflected := NOT joy.AtNeutralXY, JoystickPull := joy.AxisCmdY.DirectionPositive, JoystickPush := joy.AxisCmdY.DirectionNegative, BtnValidation := bench.Operator.JoyBtnRaw);
IF bench.Operator.JoyBtnRaw AND NOT previousButton THEN buttonEdges := buttonEdges + 1; END_IF; previousButton := bench.Operator.JoyBtnRaw;
ASSERT_FALSE(joy.DeadmanArmed, 'Pas de rearmement au retour du permis');
ADVANCE_TIME(10000000);
bench(RawPosM1 := raw1, RawPosM2 := raw2);
joy(RawX := bench.Operator.JoyXRaw_ANA1, RawY := bench.Operator.JoyYRaw_ANA2, RawButton := bench.Operator.JoyBtnRaw, Cfg := cfg, NeutralXMem := nx, NeutralYMem := ny);
home(DeadmanArmed := joy.DeadmanArmed, JoystickDeflected := NOT joy.AtNeutralXY, JoystickPull := joy.AxisCmdY.DirectionPositive, JoystickPush := joy.AxisCmdY.DirectionNegative, BtnValidation := bench.Operator.JoyBtnRaw);
IF bench.Operator.JoyBtnRaw AND NOT previousButton THEN buttonEdges := buttonEdges + 1; END_IF; previousButton := bench.Operator.JoyBtnRaw;
ASSERT_FALSE(joy.DeadmanArmed, 'Pas de rearmement au retour du permis');
ADVANCE_TIME(10000000);
bench(RawPosM1 := raw1, RawPosM2 := raw2);
joy(RawX := bench.Operator.JoyXRaw_ANA1, RawY := bench.Operator.JoyYRaw_ANA2, RawButton := bench.Operator.JoyBtnRaw, Cfg := cfg, NeutralXMem := nx, NeutralYMem := ny);
home(DeadmanArmed := joy.DeadmanArmed, JoystickDeflected := NOT joy.AtNeutralXY, JoystickPull := joy.AxisCmdY.DirectionPositive, JoystickPush := joy.AxisCmdY.DirectionNegative, BtnValidation := bench.Operator.JoyBtnRaw);
IF bench.Operator.JoyBtnRaw AND NOT previousButton THEN buttonEdges := buttonEdges + 1; END_IF; previousButton := bench.Operator.JoyBtnRaw;
ASSERT_FALSE(joy.DeadmanArmed, 'Pas de rearmement au retour du permis');
ADVANCE_TIME(10000000);
bench(RawPosM1 := raw1, RawPosM2 := raw2);
joy(RawX := bench.Operator.JoyXRaw_ANA1, RawY := bench.Operator.JoyYRaw_ANA2, RawButton := bench.Operator.JoyBtnRaw, Cfg := cfg, NeutralXMem := nx, NeutralYMem := ny);
home(DeadmanArmed := joy.DeadmanArmed, JoystickDeflected := NOT joy.AtNeutralXY, JoystickPull := joy.AxisCmdY.DirectionPositive, JoystickPush := joy.AxisCmdY.DirectionNegative, BtnValidation := bench.Operator.JoyBtnRaw);
IF bench.Operator.JoyBtnRaw AND NOT previousButton THEN buttonEdges := buttonEdges + 1; END_IF; previousButton := bench.Operator.JoyBtnRaw;
ASSERT_FALSE(joy.DeadmanArmed, 'Pas de rearmement au retour du permis');
ADVANCE_TIME(10000000);
bench(RawPosM1 := raw1, RawPosM2 := raw2);
joy(RawX := bench.Operator.JoyXRaw_ANA1, RawY := bench.Operator.JoyYRaw_ANA2, RawButton := bench.Operator.JoyBtnRaw, Cfg := cfg, NeutralXMem := nx, NeutralYMem := ny);
home(DeadmanArmed := joy.DeadmanArmed, JoystickDeflected := NOT joy.AtNeutralXY, JoystickPull := joy.AxisCmdY.DirectionPositive, JoystickPush := joy.AxisCmdY.DirectionNegative, BtnValidation := bench.Operator.JoyBtnRaw);
IF bench.Operator.JoyBtnRaw AND NOT previousButton THEN buttonEdges := buttonEdges + 1; END_IF; previousButton := bench.Operator.JoyBtnRaw;
ASSERT_FALSE(joy.DeadmanArmed, 'Pas de rearmement au retour du permis');
ADVANCE_TIME(10000000);
bench(RawPosM1 := raw1, RawPosM2 := raw2);
joy(RawX := bench.Operator.JoyXRaw_ANA1, RawY := bench.Operator.JoyYRaw_ANA2, RawButton := bench.Operator.JoyBtnRaw, Cfg := cfg, NeutralXMem := nx, NeutralYMem := ny);
home(DeadmanArmed := joy.DeadmanArmed, JoystickDeflected := NOT joy.AtNeutralXY, JoystickPull := joy.AxisCmdY.DirectionPositive, JoystickPush := joy.AxisCmdY.DirectionNegative, BtnValidation := bench.Operator.JoyBtnRaw);
IF bench.Operator.JoyBtnRaw AND NOT previousButton THEN buttonEdges := buttonEdges + 1; END_IF; previousButton := bench.Operator.JoyBtnRaw;
ASSERT_FALSE(joy.DeadmanArmed, 'Pas de rearmement au retour du permis');
ADVANCE_TIME(10000000);
bench(RawPosM1 := raw1, RawPosM2 := raw2);
joy(RawX := bench.Operator.JoyXRaw_ANA1, RawY := bench.Operator.JoyYRaw_ANA2, RawButton := bench.Operator.JoyBtnRaw, Cfg := cfg, NeutralXMem := nx, NeutralYMem := ny);
home(DeadmanArmed := joy.DeadmanArmed, JoystickDeflected := NOT joy.AtNeutralXY, JoystickPull := joy.AxisCmdY.DirectionPositive, JoystickPush := joy.AxisCmdY.DirectionNegative, BtnValidation := bench.Operator.JoyBtnRaw);
IF bench.Operator.JoyBtnRaw AND NOT previousButton THEN buttonEdges := buttonEdges + 1; END_IF; previousButton := bench.Operator.JoyBtnRaw;
ASSERT_FALSE(joy.DeadmanArmed, 'Pas de rearmement au retour du permis');
ADVANCE_TIME(10000000);
bench(RawPosM1 := raw1, RawPosM2 := raw2);
joy(RawX := bench.Operator.JoyXRaw_ANA1, RawY := bench.Operator.JoyYRaw_ANA2, RawButton := bench.Operator.JoyBtnRaw, Cfg := cfg, NeutralXMem := nx, NeutralYMem := ny);
home(DeadmanArmed := joy.DeadmanArmed, JoystickDeflected := NOT joy.AtNeutralXY, JoystickPull := joy.AxisCmdY.DirectionPositive, JoystickPush := joy.AxisCmdY.DirectionNegative, BtnValidation := bench.Operator.JoyBtnRaw);
IF bench.Operator.JoyBtnRaw AND NOT previousButton THEN buttonEdges := buttonEdges + 1; END_IF; previousButton := bench.Operator.JoyBtnRaw;
ASSERT_FALSE(joy.DeadmanArmed, 'Pas de rearmement au retour du permis');
ADVANCE_TIME(10000000);
bench(RawPosM1 := raw1, RawPosM2 := raw2);
joy(RawX := bench.Operator.JoyXRaw_ANA1, RawY := bench.Operator.JoyYRaw_ANA2, RawButton := bench.Operator.JoyBtnRaw, Cfg := cfg, NeutralXMem := nx, NeutralYMem := ny);
home(DeadmanArmed := joy.DeadmanArmed, JoystickDeflected := NOT joy.AtNeutralXY, JoystickPull := joy.AxisCmdY.DirectionPositive, JoystickPush := joy.AxisCmdY.DirectionNegative, BtnValidation := bench.Operator.JoyBtnRaw);
IF bench.Operator.JoyBtnRaw AND NOT previousButton THEN buttonEdges := buttonEdges + 1; END_IF; previousButton := bench.Operator.JoyBtnRaw;
ASSERT_FALSE(joy.DeadmanArmed, 'Pas de rearmement au retour du permis');
ADVANCE_TIME(10000000);
bench(RawPosM1 := raw1, RawPosM2 := raw2);
joy(RawX := bench.Operator.JoyXRaw_ANA1, RawY := bench.Operator.JoyYRaw_ANA2, RawButton := bench.Operator.JoyBtnRaw, Cfg := cfg, NeutralXMem := nx, NeutralYMem := ny);
home(DeadmanArmed := joy.DeadmanArmed, JoystickDeflected := NOT joy.AtNeutralXY, JoystickPull := joy.AxisCmdY.DirectionPositive, JoystickPush := joy.AxisCmdY.DirectionNegative, BtnValidation := bench.Operator.JoyBtnRaw);
IF bench.Operator.JoyBtnRaw AND NOT previousButton THEN buttonEdges := buttonEdges + 1; END_IF; previousButton := bench.Operator.JoyBtnRaw;
ASSERT_FALSE(joy.DeadmanArmed, 'Pas de rearmement au retour du permis');
ADVANCE_TIME(10000000);
bench(RawPosM1 := raw1, RawPosM2 := raw2);
joy(RawX := bench.Operator.JoyXRaw_ANA1, RawY := bench.Operator.JoyYRaw_ANA2, RawButton := bench.Operator.JoyBtnRaw, Cfg := cfg, NeutralXMem := nx, NeutralYMem := ny);
home(DeadmanArmed := joy.DeadmanArmed, JoystickDeflected := NOT joy.AtNeutralXY, JoystickPull := joy.AxisCmdY.DirectionPositive, JoystickPush := joy.AxisCmdY.DirectionNegative, BtnValidation := bench.Operator.JoyBtnRaw);
IF bench.Operator.JoyBtnRaw AND NOT previousButton THEN buttonEdges := buttonEdges + 1; END_IF; previousButton := bench.Operator.JoyBtnRaw;
ASSERT_FALSE(joy.DeadmanArmed, 'Pas de rearmement au retour du permis');
ADVANCE_TIME(10000000);
bench(RawPosM1 := raw1, RawPosM2 := raw2);
joy(RawX := bench.Operator.JoyXRaw_ANA1, RawY := bench.Operator.JoyYRaw_ANA2, RawButton := bench.Operator.JoyBtnRaw, Cfg := cfg, NeutralXMem := nx, NeutralYMem := ny);
home(DeadmanArmed := joy.DeadmanArmed, JoystickDeflected := NOT joy.AtNeutralXY, JoystickPull := joy.AxisCmdY.DirectionPositive, JoystickPush := joy.AxisCmdY.DirectionNegative, BtnValidation := bench.Operator.JoyBtnRaw);
IF bench.Operator.JoyBtnRaw AND NOT previousButton THEN buttonEdges := buttonEdges + 1; END_IF; previousButton := bench.Operator.JoyBtnRaw;
ASSERT_FALSE(joy.DeadmanArmed, 'Pas de rearmement au retour du permis');
ADVANCE_TIME(10000000);
bench(RawPosM1 := raw1, RawPosM2 := raw2);
joy(RawX := bench.Operator.JoyXRaw_ANA1, RawY := bench.Operator.JoyYRaw_ANA2, RawButton := bench.Operator.JoyBtnRaw, Cfg := cfg, NeutralXMem := nx, NeutralYMem := ny);
home(DeadmanArmed := joy.DeadmanArmed, JoystickDeflected := NOT joy.AtNeutralXY, JoystickPull := joy.AxisCmdY.DirectionPositive, JoystickPush := joy.AxisCmdY.DirectionNegative, BtnValidation := bench.Operator.JoyBtnRaw);
IF bench.Operator.JoyBtnRaw AND NOT previousButton THEN buttonEdges := buttonEdges + 1; END_IF; previousButton := bench.Operator.JoyBtnRaw;
ASSERT_FALSE(joy.DeadmanArmed, 'Pas de rearmement au retour du permis');
ADVANCE_TIME(10000000);
bench(RawPosM1 := raw1, RawPosM2 := raw2);
joy(RawX := bench.Operator.JoyXRaw_ANA1, RawY := bench.Operator.JoyYRaw_ANA2, RawButton := bench.Operator.JoyBtnRaw, Cfg := cfg, NeutralXMem := nx, NeutralYMem := ny);
home(DeadmanArmed := joy.DeadmanArmed, JoystickDeflected := NOT joy.AtNeutralXY, JoystickPull := joy.AxisCmdY.DirectionPositive, JoystickPush := joy.AxisCmdY.DirectionNegative, BtnValidation := bench.Operator.JoyBtnRaw);
IF bench.Operator.JoyBtnRaw AND NOT previousButton THEN buttonEdges := buttonEdges + 1; END_IF; previousButton := bench.Operator.JoyBtnRaw;
ASSERT_FALSE(joy.DeadmanArmed, 'Pas de rearmement au retour du permis');
ADVANCE_TIME(10000000);
bench(RawPosM1 := raw1, RawPosM2 := raw2);
joy(RawX := bench.Operator.JoyXRaw_ANA1, RawY := bench.Operator.JoyYRaw_ANA2, RawButton := bench.Operator.JoyBtnRaw, Cfg := cfg, NeutralXMem := nx, NeutralYMem := ny);
home(DeadmanArmed := joy.DeadmanArmed, JoystickDeflected := NOT joy.AtNeutralXY, JoystickPull := joy.AxisCmdY.DirectionPositive, JoystickPush := joy.AxisCmdY.DirectionNegative, BtnValidation := bench.Operator.JoyBtnRaw);
IF bench.Operator.JoyBtnRaw AND NOT previousButton THEN buttonEdges := buttonEdges + 1; END_IF; previousButton := bench.Operator.JoyBtnRaw;
ASSERT_FALSE(joy.DeadmanArmed, 'Pas de rearmement au retour du permis');
ADVANCE_TIME(10000000);
bench(RawPosM1 := raw1, RawPosM2 := raw2);
joy(RawX := bench.Operator.JoyXRaw_ANA1, RawY := bench.Operator.JoyYRaw_ANA2, RawButton := bench.Operator.JoyBtnRaw, Cfg := cfg, NeutralXMem := nx, NeutralYMem := ny);
home(DeadmanArmed := joy.DeadmanArmed, JoystickDeflected := NOT joy.AtNeutralXY, JoystickPull := joy.AxisCmdY.DirectionPositive, JoystickPush := joy.AxisCmdY.DirectionNegative, BtnValidation := bench.Operator.JoyBtnRaw);
IF bench.Operator.JoyBtnRaw AND NOT previousButton THEN buttonEdges := buttonEdges + 1; END_IF; previousButton := bench.Operator.JoyBtnRaw;
ASSERT_FALSE(joy.DeadmanArmed, 'Pas de rearmement au retour du permis');
ADVANCE_TIME(10000000);
bench(RawPosM1 := raw1, RawPosM2 := raw2);
joy(RawX := bench.Operator.JoyXRaw_ANA1, RawY := bench.Operator.JoyYRaw_ANA2, RawButton := bench.Operator.JoyBtnRaw, Cfg := cfg, NeutralXMem := nx, NeutralYMem := ny);
home(DeadmanArmed := joy.DeadmanArmed, JoystickDeflected := NOT joy.AtNeutralXY, JoystickPull := joy.AxisCmdY.DirectionPositive, JoystickPush := joy.AxisCmdY.DirectionNegative, BtnValidation := bench.Operator.JoyBtnRaw);
IF bench.Operator.JoyBtnRaw AND NOT previousButton THEN buttonEdges := buttonEdges + 1; END_IF; previousButton := bench.Operator.JoyBtnRaw;
ASSERT_FALSE(joy.DeadmanArmed, 'Pas de rearmement au retour du permis');
ADVANCE_TIME(10000000);
bench(RawPosM1 := raw1, RawPosM2 := raw2);
joy(RawX := bench.Operator.JoyXRaw_ANA1, RawY := bench.Operator.JoyYRaw_ANA2, RawButton := bench.Operator.JoyBtnRaw, Cfg := cfg, NeutralXMem := nx, NeutralYMem := ny);
home(DeadmanArmed := joy.DeadmanArmed, JoystickDeflected := NOT joy.AtNeutralXY, JoystickPull := joy.AxisCmdY.DirectionPositive, JoystickPush := joy.AxisCmdY.DirectionNegative, BtnValidation := bench.Operator.JoyBtnRaw);
IF bench.Operator.JoyBtnRaw AND NOT previousButton THEN buttonEdges := buttonEdges + 1; END_IF; previousButton := bench.Operator.JoyBtnRaw;
ASSERT_FALSE(joy.DeadmanArmed, 'Pas de rearmement au retour du permis');
ADVANCE_TIME(10000000);
bench(RawPosM1 := raw1, RawPosM2 := raw2);
joy(RawX := bench.Operator.JoyXRaw_ANA1, RawY := bench.Operator.JoyYRaw_ANA2, RawButton := bench.Operator.JoyBtnRaw, Cfg := cfg, NeutralXMem := nx, NeutralYMem := ny);
home(DeadmanArmed := joy.DeadmanArmed, JoystickDeflected := NOT joy.AtNeutralXY, JoystickPull := joy.AxisCmdY.DirectionPositive, JoystickPush := joy.AxisCmdY.DirectionNegative, BtnValidation := bench.Operator.JoyBtnRaw);
IF bench.Operator.JoyBtnRaw AND NOT previousButton THEN buttonEdges := buttonEdges + 1; END_IF; previousButton := bench.Operator.JoyBtnRaw;
ASSERT_FALSE(joy.DeadmanArmed, 'Pas de rearmement au retour du permis');
ADVANCE_TIME(10000000);
bench(RawPosM1 := raw1, RawPosM2 := raw2);
joy(RawX := bench.Operator.JoyXRaw_ANA1, RawY := bench.Operator.JoyYRaw_ANA2, RawButton := bench.Operator.JoyBtnRaw, Cfg := cfg, NeutralXMem := nx, NeutralYMem := ny);
home(DeadmanArmed := joy.DeadmanArmed, JoystickDeflected := NOT joy.AtNeutralXY, JoystickPull := joy.AxisCmdY.DirectionPositive, JoystickPush := joy.AxisCmdY.DirectionNegative, BtnValidation := bench.Operator.JoyBtnRaw);
IF bench.Operator.JoyBtnRaw AND NOT previousButton THEN buttonEdges := buttonEdges + 1; END_IF; previousButton := bench.Operator.JoyBtnRaw;
ASSERT_FALSE(joy.DeadmanArmed, 'Pas de rearmement au retour du permis');
ADVANCE_TIME(10000000);
bench(RawPosM1 := raw1, RawPosM2 := raw2);
joy(RawX := bench.Operator.JoyXRaw_ANA1, RawY := bench.Operator.JoyYRaw_ANA2, RawButton := bench.Operator.JoyBtnRaw, Cfg := cfg, NeutralXMem := nx, NeutralYMem := ny);
home(DeadmanArmed := joy.DeadmanArmed, JoystickDeflected := NOT joy.AtNeutralXY, JoystickPull := joy.AxisCmdY.DirectionPositive, JoystickPush := joy.AxisCmdY.DirectionNegative, BtnValidation := bench.Operator.JoyBtnRaw);
IF bench.Operator.JoyBtnRaw AND NOT previousButton THEN buttonEdges := buttonEdges + 1; END_IF; previousButton := bench.Operator.JoyBtnRaw;
ASSERT_FALSE(joy.DeadmanArmed, 'Pas de rearmement au retour du permis');
ADVANCE_TIME(10000000);
bench(RawPosM1 := raw1, RawPosM2 := raw2);
joy(RawX := bench.Operator.JoyXRaw_ANA1, RawY := bench.Operator.JoyYRaw_ANA2, RawButton := bench.Operator.JoyBtnRaw, Cfg := cfg, NeutralXMem := nx, NeutralYMem := ny);
home(DeadmanArmed := joy.DeadmanArmed, JoystickDeflected := NOT joy.AtNeutralXY, JoystickPull := joy.AxisCmdY.DirectionPositive, JoystickPush := joy.AxisCmdY.DirectionNegative, BtnValidation := bench.Operator.JoyBtnRaw);
IF bench.Operator.JoyBtnRaw AND NOT previousButton THEN buttonEdges := buttonEdges + 1; END_IF; previousButton := bench.Operator.JoyBtnRaw;
ASSERT_FALSE(joy.DeadmanArmed, 'Pas de rearmement au retour du permis');
ADVANCE_TIME(10000000);
bench(RawPosM1 := raw1, RawPosM2 := raw2);
joy(RawX := bench.Operator.JoyXRaw_ANA1, RawY := bench.Operator.JoyYRaw_ANA2, RawButton := bench.Operator.JoyBtnRaw, Cfg := cfg, NeutralXMem := nx, NeutralYMem := ny);
home(DeadmanArmed := joy.DeadmanArmed, JoystickDeflected := NOT joy.AtNeutralXY, JoystickPull := joy.AxisCmdY.DirectionPositive, JoystickPush := joy.AxisCmdY.DirectionNegative, BtnValidation := bench.Operator.JoyBtnRaw);
IF bench.Operator.JoyBtnRaw AND NOT previousButton THEN buttonEdges := buttonEdges + 1; END_IF; previousButton := bench.Operator.JoyBtnRaw;
ASSERT_FALSE(joy.DeadmanArmed, 'Pas de rearmement au retour du permis');
ASSERT_EQ(buttonEdges, 1, 'Aucune nouvelle tentative');
END_TEST

TEST 'TC-T418-INT-003 Perte permis pendant geste arme'
nx := 5000; ny := 5000; raw1 := 0; raw2 := 0; previousButton := FALSE; buttonEdges := 0;
bench.Enable := TRUE; joy.Enable := TRUE; joy.ArmingPermit := TRUE; diagOk.Operational := TRUE;
joy.BusCanOpenOP := diagOk; joy.JoystickOP := diagOk; home.Enable := TRUE; home.BootReady := TRUE;
home.Mode := E_Mode.MAINT_N1; home.BucketOffsetValid := TRUE; home.WinchesMechanicallyStopped := TRUE;
ADVANCE_TIME(10000000);
bench(RawPosM1 := raw1, RawPosM2 := raw2);
joy(RawX := bench.Operator.JoyXRaw_ANA1, RawY := bench.Operator.JoyYRaw_ANA2, RawButton := bench.Operator.JoyBtnRaw, Cfg := cfg, NeutralXMem := nx, NeutralYMem := ny);
home(DeadmanArmed := joy.DeadmanArmed, JoystickDeflected := NOT joy.AtNeutralXY, JoystickPull := joy.AxisCmdY.DirectionPositive, JoystickPush := joy.AxisCmdY.DirectionNegative, BtnValidation := bench.Operator.JoyBtnRaw);
IF bench.Operator.JoyBtnRaw AND NOT previousButton THEN buttonEdges := buttonEdges + 1; END_IF; previousButton := bench.Operator.JoyBtnRaw;
bench.SimJoystickRev_Down_Open_Active := TRUE;
ADVANCE_TIME(10000000);
bench(RawPosM1 := raw1, RawPosM2 := raw2);
joy(RawX := bench.Operator.JoyXRaw_ANA1, RawY := bench.Operator.JoyYRaw_ANA2, RawButton := bench.Operator.JoyBtnRaw, Cfg := cfg, NeutralXMem := nx, NeutralYMem := ny);
home(DeadmanArmed := joy.DeadmanArmed, JoystickDeflected := NOT joy.AtNeutralXY, JoystickPull := joy.AxisCmdY.DirectionPositive, JoystickPush := joy.AxisCmdY.DirectionNegative, BtnValidation := bench.Operator.JoyBtnRaw);
IF bench.Operator.JoyBtnRaw AND NOT previousButton THEN buttonEdges := buttonEdges + 1; END_IF; previousButton := bench.Operator.JoyBtnRaw;
ADVANCE_TIME(10000000);
bench(RawPosM1 := raw1, RawPosM2 := raw2);
joy(RawX := bench.Operator.JoyXRaw_ANA1, RawY := bench.Operator.JoyYRaw_ANA2, RawButton := bench.Operator.JoyBtnRaw, Cfg := cfg, NeutralXMem := nx, NeutralYMem := ny);
home(DeadmanArmed := joy.DeadmanArmed, JoystickDeflected := NOT joy.AtNeutralXY, JoystickPull := joy.AxisCmdY.DirectionPositive, JoystickPush := joy.AxisCmdY.DirectionNegative, BtnValidation := bench.Operator.JoyBtnRaw);
IF bench.Operator.JoyBtnRaw AND NOT previousButton THEN buttonEdges := buttonEdges + 1; END_IF; previousButton := bench.Operator.JoyBtnRaw;
ADVANCE_TIME(10000000);
bench(RawPosM1 := raw1, RawPosM2 := raw2);
joy(RawX := bench.Operator.JoyXRaw_ANA1, RawY := bench.Operator.JoyYRaw_ANA2, RawButton := bench.Operator.JoyBtnRaw, Cfg := cfg, NeutralXMem := nx, NeutralYMem := ny);
home(DeadmanArmed := joy.DeadmanArmed, JoystickDeflected := NOT joy.AtNeutralXY, JoystickPull := joy.AxisCmdY.DirectionPositive, JoystickPush := joy.AxisCmdY.DirectionNegative, BtnValidation := bench.Operator.JoyBtnRaw);
IF bench.Operator.JoyBtnRaw AND NOT previousButton THEN buttonEdges := buttonEdges + 1; END_IF; previousButton := bench.Operator.JoyBtnRaw;
ADVANCE_TIME(10000000);
bench(RawPosM1 := raw1, RawPosM2 := raw2);
joy(RawX := bench.Operator.JoyXRaw_ANA1, RawY := bench.Operator.JoyYRaw_ANA2, RawButton := bench.Operator.JoyBtnRaw, Cfg := cfg, NeutralXMem := nx, NeutralYMem := ny);
home(DeadmanArmed := joy.DeadmanArmed, JoystickDeflected := NOT joy.AtNeutralXY, JoystickPull := joy.AxisCmdY.DirectionPositive, JoystickPush := joy.AxisCmdY.DirectionNegative, BtnValidation := bench.Operator.JoyBtnRaw);
IF bench.Operator.JoyBtnRaw AND NOT previousButton THEN buttonEdges := buttonEdges + 1; END_IF; previousButton := bench.Operator.JoyBtnRaw;
ADVANCE_TIME(10000000);
bench(RawPosM1 := raw1, RawPosM2 := raw2);
joy(RawX := bench.Operator.JoyXRaw_ANA1, RawY := bench.Operator.JoyYRaw_ANA2, RawButton := bench.Operator.JoyBtnRaw, Cfg := cfg, NeutralXMem := nx, NeutralYMem := ny);
home(DeadmanArmed := joy.DeadmanArmed, JoystickDeflected := NOT joy.AtNeutralXY, JoystickPull := joy.AxisCmdY.DirectionPositive, JoystickPush := joy.AxisCmdY.DirectionNegative, BtnValidation := bench.Operator.JoyBtnRaw);
IF bench.Operator.JoyBtnRaw AND NOT previousButton THEN buttonEdges := buttonEdges + 1; END_IF; previousButton := bench.Operator.JoyBtnRaw;
ADVANCE_TIME(10000000);
bench(RawPosM1 := raw1, RawPosM2 := raw2);
joy(RawX := bench.Operator.JoyXRaw_ANA1, RawY := bench.Operator.JoyYRaw_ANA2, RawButton := bench.Operator.JoyBtnRaw, Cfg := cfg, NeutralXMem := nx, NeutralYMem := ny);
home(DeadmanArmed := joy.DeadmanArmed, JoystickDeflected := NOT joy.AtNeutralXY, JoystickPull := joy.AxisCmdY.DirectionPositive, JoystickPush := joy.AxisCmdY.DirectionNegative, BtnValidation := bench.Operator.JoyBtnRaw);
IF bench.Operator.JoyBtnRaw AND NOT previousButton THEN buttonEdges := buttonEdges + 1; END_IF; previousButton := bench.Operator.JoyBtnRaw;
ADVANCE_TIME(10000000);
bench(RawPosM1 := raw1, RawPosM2 := raw2);
joy(RawX := bench.Operator.JoyXRaw_ANA1, RawY := bench.Operator.JoyYRaw_ANA2, RawButton := bench.Operator.JoyBtnRaw, Cfg := cfg, NeutralXMem := nx, NeutralYMem := ny);
home(DeadmanArmed := joy.DeadmanArmed, JoystickDeflected := NOT joy.AtNeutralXY, JoystickPull := joy.AxisCmdY.DirectionPositive, JoystickPush := joy.AxisCmdY.DirectionNegative, BtnValidation := bench.Operator.JoyBtnRaw);
IF bench.Operator.JoyBtnRaw AND NOT previousButton THEN buttonEdges := buttonEdges + 1; END_IF; previousButton := bench.Operator.JoyBtnRaw;
ADVANCE_TIME(10000000);
bench(RawPosM1 := raw1, RawPosM2 := raw2);
joy(RawX := bench.Operator.JoyXRaw_ANA1, RawY := bench.Operator.JoyYRaw_ANA2, RawButton := bench.Operator.JoyBtnRaw, Cfg := cfg, NeutralXMem := nx, NeutralYMem := ny);
home(DeadmanArmed := joy.DeadmanArmed, JoystickDeflected := NOT joy.AtNeutralXY, JoystickPull := joy.AxisCmdY.DirectionPositive, JoystickPush := joy.AxisCmdY.DirectionNegative, BtnValidation := bench.Operator.JoyBtnRaw);
IF bench.Operator.JoyBtnRaw AND NOT previousButton THEN buttonEdges := buttonEdges + 1; END_IF; previousButton := bench.Operator.JoyBtnRaw;
ADVANCE_TIME(10000000);
bench(RawPosM1 := raw1, RawPosM2 := raw2);
joy(RawX := bench.Operator.JoyXRaw_ANA1, RawY := bench.Operator.JoyYRaw_ANA2, RawButton := bench.Operator.JoyBtnRaw, Cfg := cfg, NeutralXMem := nx, NeutralYMem := ny);
home(DeadmanArmed := joy.DeadmanArmed, JoystickDeflected := NOT joy.AtNeutralXY, JoystickPull := joy.AxisCmdY.DirectionPositive, JoystickPush := joy.AxisCmdY.DirectionNegative, BtnValidation := bench.Operator.JoyBtnRaw);
IF bench.Operator.JoyBtnRaw AND NOT previousButton THEN buttonEdges := buttonEdges + 1; END_IF; previousButton := bench.Operator.JoyBtnRaw;
ADVANCE_TIME(10000000);
bench(RawPosM1 := raw1, RawPosM2 := raw2);
joy(RawX := bench.Operator.JoyXRaw_ANA1, RawY := bench.Operator.JoyYRaw_ANA2, RawButton := bench.Operator.JoyBtnRaw, Cfg := cfg, NeutralXMem := nx, NeutralYMem := ny);
home(DeadmanArmed := joy.DeadmanArmed, JoystickDeflected := NOT joy.AtNeutralXY, JoystickPull := joy.AxisCmdY.DirectionPositive, JoystickPush := joy.AxisCmdY.DirectionNegative, BtnValidation := bench.Operator.JoyBtnRaw);
IF bench.Operator.JoyBtnRaw AND NOT previousButton THEN buttonEdges := buttonEdges + 1; END_IF; previousButton := bench.Operator.JoyBtnRaw;
ADVANCE_TIME(10000000);
bench(RawPosM1 := raw1, RawPosM2 := raw2);
joy(RawX := bench.Operator.JoyXRaw_ANA1, RawY := bench.Operator.JoyYRaw_ANA2, RawButton := bench.Operator.JoyBtnRaw, Cfg := cfg, NeutralXMem := nx, NeutralYMem := ny);
home(DeadmanArmed := joy.DeadmanArmed, JoystickDeflected := NOT joy.AtNeutralXY, JoystickPull := joy.AxisCmdY.DirectionPositive, JoystickPush := joy.AxisCmdY.DirectionNegative, BtnValidation := bench.Operator.JoyBtnRaw);
IF bench.Operator.JoyBtnRaw AND NOT previousButton THEN buttonEdges := buttonEdges + 1; END_IF; previousButton := bench.Operator.JoyBtnRaw;
ADVANCE_TIME(10000000);
bench(RawPosM1 := raw1, RawPosM2 := raw2);
joy(RawX := bench.Operator.JoyXRaw_ANA1, RawY := bench.Operator.JoyYRaw_ANA2, RawButton := bench.Operator.JoyBtnRaw, Cfg := cfg, NeutralXMem := nx, NeutralYMem := ny);
home(DeadmanArmed := joy.DeadmanArmed, JoystickDeflected := NOT joy.AtNeutralXY, JoystickPull := joy.AxisCmdY.DirectionPositive, JoystickPush := joy.AxisCmdY.DirectionNegative, BtnValidation := bench.Operator.JoyBtnRaw);
IF bench.Operator.JoyBtnRaw AND NOT previousButton THEN buttonEdges := buttonEdges + 1; END_IF; previousButton := bench.Operator.JoyBtnRaw;
ADVANCE_TIME(10000000);
bench(RawPosM1 := raw1, RawPosM2 := raw2);
joy(RawX := bench.Operator.JoyXRaw_ANA1, RawY := bench.Operator.JoyYRaw_ANA2, RawButton := bench.Operator.JoyBtnRaw, Cfg := cfg, NeutralXMem := nx, NeutralYMem := ny);
home(DeadmanArmed := joy.DeadmanArmed, JoystickDeflected := NOT joy.AtNeutralXY, JoystickPull := joy.AxisCmdY.DirectionPositive, JoystickPush := joy.AxisCmdY.DirectionNegative, BtnValidation := bench.Operator.JoyBtnRaw);
IF bench.Operator.JoyBtnRaw AND NOT previousButton THEN buttonEdges := buttonEdges + 1; END_IF; previousButton := bench.Operator.JoyBtnRaw;
ADVANCE_TIME(10000000);
bench(RawPosM1 := raw1, RawPosM2 := raw2);
joy(RawX := bench.Operator.JoyXRaw_ANA1, RawY := bench.Operator.JoyYRaw_ANA2, RawButton := bench.Operator.JoyBtnRaw, Cfg := cfg, NeutralXMem := nx, NeutralYMem := ny);
home(DeadmanArmed := joy.DeadmanArmed, JoystickDeflected := NOT joy.AtNeutralXY, JoystickPull := joy.AxisCmdY.DirectionPositive, JoystickPush := joy.AxisCmdY.DirectionNegative, BtnValidation := bench.Operator.JoyBtnRaw);
IF bench.Operator.JoyBtnRaw AND NOT previousButton THEN buttonEdges := buttonEdges + 1; END_IF; previousButton := bench.Operator.JoyBtnRaw;
ADVANCE_TIME(10000000);
bench(RawPosM1 := raw1, RawPosM2 := raw2);
joy(RawX := bench.Operator.JoyXRaw_ANA1, RawY := bench.Operator.JoyYRaw_ANA2, RawButton := bench.Operator.JoyBtnRaw, Cfg := cfg, NeutralXMem := nx, NeutralYMem := ny);
home(DeadmanArmed := joy.DeadmanArmed, JoystickDeflected := NOT joy.AtNeutralXY, JoystickPull := joy.AxisCmdY.DirectionPositive, JoystickPush := joy.AxisCmdY.DirectionNegative, BtnValidation := bench.Operator.JoyBtnRaw);
IF bench.Operator.JoyBtnRaw AND NOT previousButton THEN buttonEdges := buttonEdges + 1; END_IF; previousButton := bench.Operator.JoyBtnRaw;
ADVANCE_TIME(10000000);
bench(RawPosM1 := raw1, RawPosM2 := raw2);
joy(RawX := bench.Operator.JoyXRaw_ANA1, RawY := bench.Operator.JoyYRaw_ANA2, RawButton := bench.Operator.JoyBtnRaw, Cfg := cfg, NeutralXMem := nx, NeutralYMem := ny);
home(DeadmanArmed := joy.DeadmanArmed, JoystickDeflected := NOT joy.AtNeutralXY, JoystickPull := joy.AxisCmdY.DirectionPositive, JoystickPush := joy.AxisCmdY.DirectionNegative, BtnValidation := bench.Operator.JoyBtnRaw);
IF bench.Operator.JoyBtnRaw AND NOT previousButton THEN buttonEdges := buttonEdges + 1; END_IF; previousButton := bench.Operator.JoyBtnRaw;
ADVANCE_TIME(10000000);
bench(RawPosM1 := raw1, RawPosM2 := raw2);
joy(RawX := bench.Operator.JoyXRaw_ANA1, RawY := bench.Operator.JoyYRaw_ANA2, RawButton := bench.Operator.JoyBtnRaw, Cfg := cfg, NeutralXMem := nx, NeutralYMem := ny);
home(DeadmanArmed := joy.DeadmanArmed, JoystickDeflected := NOT joy.AtNeutralXY, JoystickPull := joy.AxisCmdY.DirectionPositive, JoystickPush := joy.AxisCmdY.DirectionNegative, BtnValidation := bench.Operator.JoyBtnRaw);
IF bench.Operator.JoyBtnRaw AND NOT previousButton THEN buttonEdges := buttonEdges + 1; END_IF; previousButton := bench.Operator.JoyBtnRaw;
ADVANCE_TIME(10000000);
bench(RawPosM1 := raw1, RawPosM2 := raw2);
joy(RawX := bench.Operator.JoyXRaw_ANA1, RawY := bench.Operator.JoyYRaw_ANA2, RawButton := bench.Operator.JoyBtnRaw, Cfg := cfg, NeutralXMem := nx, NeutralYMem := ny);
home(DeadmanArmed := joy.DeadmanArmed, JoystickDeflected := NOT joy.AtNeutralXY, JoystickPull := joy.AxisCmdY.DirectionPositive, JoystickPush := joy.AxisCmdY.DirectionNegative, BtnValidation := bench.Operator.JoyBtnRaw);
IF bench.Operator.JoyBtnRaw AND NOT previousButton THEN buttonEdges := buttonEdges + 1; END_IF; previousButton := bench.Operator.JoyBtnRaw;
ADVANCE_TIME(10000000);
bench(RawPosM1 := raw1, RawPosM2 := raw2);
joy(RawX := bench.Operator.JoyXRaw_ANA1, RawY := bench.Operator.JoyYRaw_ANA2, RawButton := bench.Operator.JoyBtnRaw, Cfg := cfg, NeutralXMem := nx, NeutralYMem := ny);
home(DeadmanArmed := joy.DeadmanArmed, JoystickDeflected := NOT joy.AtNeutralXY, JoystickPull := joy.AxisCmdY.DirectionPositive, JoystickPush := joy.AxisCmdY.DirectionNegative, BtnValidation := bench.Operator.JoyBtnRaw);
IF bench.Operator.JoyBtnRaw AND NOT previousButton THEN buttonEdges := buttonEdges + 1; END_IF; previousButton := bench.Operator.JoyBtnRaw;
ADVANCE_TIME(10000000);
bench(RawPosM1 := raw1, RawPosM2 := raw2);
joy(RawX := bench.Operator.JoyXRaw_ANA1, RawY := bench.Operator.JoyYRaw_ANA2, RawButton := bench.Operator.JoyBtnRaw, Cfg := cfg, NeutralXMem := nx, NeutralYMem := ny);
home(DeadmanArmed := joy.DeadmanArmed, JoystickDeflected := NOT joy.AtNeutralXY, JoystickPull := joy.AxisCmdY.DirectionPositive, JoystickPush := joy.AxisCmdY.DirectionNegative, BtnValidation := bench.Operator.JoyBtnRaw);
IF bench.Operator.JoyBtnRaw AND NOT previousButton THEN buttonEdges := buttonEdges + 1; END_IF; previousButton := bench.Operator.JoyBtnRaw;
ADVANCE_TIME(10000000);
bench(RawPosM1 := raw1, RawPosM2 := raw2);
joy(RawX := bench.Operator.JoyXRaw_ANA1, RawY := bench.Operator.JoyYRaw_ANA2, RawButton := bench.Operator.JoyBtnRaw, Cfg := cfg, NeutralXMem := nx, NeutralYMem := ny);
home(DeadmanArmed := joy.DeadmanArmed, JoystickDeflected := NOT joy.AtNeutralXY, JoystickPull := joy.AxisCmdY.DirectionPositive, JoystickPush := joy.AxisCmdY.DirectionNegative, BtnValidation := bench.Operator.JoyBtnRaw);
IF bench.Operator.JoyBtnRaw AND NOT previousButton THEN buttonEdges := buttonEdges + 1; END_IF; previousButton := bench.Operator.JoyBtnRaw;
ADVANCE_TIME(10000000);
bench(RawPosM1 := raw1, RawPosM2 := raw2);
joy(RawX := bench.Operator.JoyXRaw_ANA1, RawY := bench.Operator.JoyYRaw_ANA2, RawButton := bench.Operator.JoyBtnRaw, Cfg := cfg, NeutralXMem := nx, NeutralYMem := ny);
home(DeadmanArmed := joy.DeadmanArmed, JoystickDeflected := NOT joy.AtNeutralXY, JoystickPull := joy.AxisCmdY.DirectionPositive, JoystickPush := joy.AxisCmdY.DirectionNegative, BtnValidation := bench.Operator.JoyBtnRaw);
IF bench.Operator.JoyBtnRaw AND NOT previousButton THEN buttonEdges := buttonEdges + 1; END_IF; previousButton := bench.Operator.JoyBtnRaw;
ADVANCE_TIME(10000000);
bench(RawPosM1 := raw1, RawPosM2 := raw2);
joy(RawX := bench.Operator.JoyXRaw_ANA1, RawY := bench.Operator.JoyYRaw_ANA2, RawButton := bench.Operator.JoyBtnRaw, Cfg := cfg, NeutralXMem := nx, NeutralYMem := ny);
home(DeadmanArmed := joy.DeadmanArmed, JoystickDeflected := NOT joy.AtNeutralXY, JoystickPull := joy.AxisCmdY.DirectionPositive, JoystickPush := joy.AxisCmdY.DirectionNegative, BtnValidation := bench.Operator.JoyBtnRaw);
IF bench.Operator.JoyBtnRaw AND NOT previousButton THEN buttonEdges := buttonEdges + 1; END_IF; previousButton := bench.Operator.JoyBtnRaw;
ADVANCE_TIME(10000000);
bench(RawPosM1 := raw1, RawPosM2 := raw2);
joy(RawX := bench.Operator.JoyXRaw_ANA1, RawY := bench.Operator.JoyYRaw_ANA2, RawButton := bench.Operator.JoyBtnRaw, Cfg := cfg, NeutralXMem := nx, NeutralYMem := ny);
home(DeadmanArmed := joy.DeadmanArmed, JoystickDeflected := NOT joy.AtNeutralXY, JoystickPull := joy.AxisCmdY.DirectionPositive, JoystickPush := joy.AxisCmdY.DirectionNegative, BtnValidation := bench.Operator.JoyBtnRaw);
IF bench.Operator.JoyBtnRaw AND NOT previousButton THEN buttonEdges := buttonEdges + 1; END_IF; previousButton := bench.Operator.JoyBtnRaw;
ADVANCE_TIME(10000000);
bench(RawPosM1 := raw1, RawPosM2 := raw2);
joy(RawX := bench.Operator.JoyXRaw_ANA1, RawY := bench.Operator.JoyYRaw_ANA2, RawButton := bench.Operator.JoyBtnRaw, Cfg := cfg, NeutralXMem := nx, NeutralYMem := ny);
home(DeadmanArmed := joy.DeadmanArmed, JoystickDeflected := NOT joy.AtNeutralXY, JoystickPull := joy.AxisCmdY.DirectionPositive, JoystickPush := joy.AxisCmdY.DirectionNegative, BtnValidation := bench.Operator.JoyBtnRaw);
IF bench.Operator.JoyBtnRaw AND NOT previousButton THEN buttonEdges := buttonEdges + 1; END_IF; previousButton := bench.Operator.JoyBtnRaw;
ADVANCE_TIME(10000000);
bench(RawPosM1 := raw1, RawPosM2 := raw2);
joy(RawX := bench.Operator.JoyXRaw_ANA1, RawY := bench.Operator.JoyYRaw_ANA2, RawButton := bench.Operator.JoyBtnRaw, Cfg := cfg, NeutralXMem := nx, NeutralYMem := ny);
home(DeadmanArmed := joy.DeadmanArmed, JoystickDeflected := NOT joy.AtNeutralXY, JoystickPull := joy.AxisCmdY.DirectionPositive, JoystickPush := joy.AxisCmdY.DirectionNegative, BtnValidation := bench.Operator.JoyBtnRaw);
IF bench.Operator.JoyBtnRaw AND NOT previousButton THEN buttonEdges := buttonEdges + 1; END_IF; previousButton := bench.Operator.JoyBtnRaw;
ADVANCE_TIME(10000000);
bench(RawPosM1 := raw1, RawPosM2 := raw2);
joy(RawX := bench.Operator.JoyXRaw_ANA1, RawY := bench.Operator.JoyYRaw_ANA2, RawButton := bench.Operator.JoyBtnRaw, Cfg := cfg, NeutralXMem := nx, NeutralYMem := ny);
home(DeadmanArmed := joy.DeadmanArmed, JoystickDeflected := NOT joy.AtNeutralXY, JoystickPull := joy.AxisCmdY.DirectionPositive, JoystickPush := joy.AxisCmdY.DirectionNegative, BtnValidation := bench.Operator.JoyBtnRaw);
IF bench.Operator.JoyBtnRaw AND NOT previousButton THEN buttonEdges := buttonEdges + 1; END_IF; previousButton := bench.Operator.JoyBtnRaw;
ADVANCE_TIME(10000000);
bench(RawPosM1 := raw1, RawPosM2 := raw2);
joy(RawX := bench.Operator.JoyXRaw_ANA1, RawY := bench.Operator.JoyYRaw_ANA2, RawButton := bench.Operator.JoyBtnRaw, Cfg := cfg, NeutralXMem := nx, NeutralYMem := ny);
home(DeadmanArmed := joy.DeadmanArmed, JoystickDeflected := NOT joy.AtNeutralXY, JoystickPull := joy.AxisCmdY.DirectionPositive, JoystickPush := joy.AxisCmdY.DirectionNegative, BtnValidation := bench.Operator.JoyBtnRaw);
IF bench.Operator.JoyBtnRaw AND NOT previousButton THEN buttonEdges := buttonEdges + 1; END_IF; previousButton := bench.Operator.JoyBtnRaw;
ADVANCE_TIME(10000000);
bench(RawPosM1 := raw1, RawPosM2 := raw2);
joy(RawX := bench.Operator.JoyXRaw_ANA1, RawY := bench.Operator.JoyYRaw_ANA2, RawButton := bench.Operator.JoyBtnRaw, Cfg := cfg, NeutralXMem := nx, NeutralYMem := ny);
home(DeadmanArmed := joy.DeadmanArmed, JoystickDeflected := NOT joy.AtNeutralXY, JoystickPull := joy.AxisCmdY.DirectionPositive, JoystickPush := joy.AxisCmdY.DirectionNegative, BtnValidation := bench.Operator.JoyBtnRaw);
IF bench.Operator.JoyBtnRaw AND NOT previousButton THEN buttonEdges := buttonEdges + 1; END_IF; previousButton := bench.Operator.JoyBtnRaw;
ADVANCE_TIME(10000000);
bench(RawPosM1 := raw1, RawPosM2 := raw2);
joy(RawX := bench.Operator.JoyXRaw_ANA1, RawY := bench.Operator.JoyYRaw_ANA2, RawButton := bench.Operator.JoyBtnRaw, Cfg := cfg, NeutralXMem := nx, NeutralYMem := ny);
home(DeadmanArmed := joy.DeadmanArmed, JoystickDeflected := NOT joy.AtNeutralXY, JoystickPull := joy.AxisCmdY.DirectionPositive, JoystickPush := joy.AxisCmdY.DirectionNegative, BtnValidation := bench.Operator.JoyBtnRaw);
IF bench.Operator.JoyBtnRaw AND NOT previousButton THEN buttonEdges := buttonEdges + 1; END_IF; previousButton := bench.Operator.JoyBtnRaw;
ADVANCE_TIME(10000000);
bench(RawPosM1 := raw1, RawPosM2 := raw2);
joy(RawX := bench.Operator.JoyXRaw_ANA1, RawY := bench.Operator.JoyYRaw_ANA2, RawButton := bench.Operator.JoyBtnRaw, Cfg := cfg, NeutralXMem := nx, NeutralYMem := ny);
home(DeadmanArmed := joy.DeadmanArmed, JoystickDeflected := NOT joy.AtNeutralXY, JoystickPull := joy.AxisCmdY.DirectionPositive, JoystickPush := joy.AxisCmdY.DirectionNegative, BtnValidation := bench.Operator.JoyBtnRaw);
IF bench.Operator.JoyBtnRaw AND NOT previousButton THEN buttonEdges := buttonEdges + 1; END_IF; previousButton := bench.Operator.JoyBtnRaw;
ADVANCE_TIME(10000000);
bench(RawPosM1 := raw1, RawPosM2 := raw2);
joy(RawX := bench.Operator.JoyXRaw_ANA1, RawY := bench.Operator.JoyYRaw_ANA2, RawButton := bench.Operator.JoyBtnRaw, Cfg := cfg, NeutralXMem := nx, NeutralYMem := ny);
home(DeadmanArmed := joy.DeadmanArmed, JoystickDeflected := NOT joy.AtNeutralXY, JoystickPull := joy.AxisCmdY.DirectionPositive, JoystickPush := joy.AxisCmdY.DirectionNegative, BtnValidation := bench.Operator.JoyBtnRaw);
IF bench.Operator.JoyBtnRaw AND NOT previousButton THEN buttonEdges := buttonEdges + 1; END_IF; previousButton := bench.Operator.JoyBtnRaw;
ADVANCE_TIME(10000000);
bench(RawPosM1 := raw1, RawPosM2 := raw2);
joy(RawX := bench.Operator.JoyXRaw_ANA1, RawY := bench.Operator.JoyYRaw_ANA2, RawButton := bench.Operator.JoyBtnRaw, Cfg := cfg, NeutralXMem := nx, NeutralYMem := ny);
home(DeadmanArmed := joy.DeadmanArmed, JoystickDeflected := NOT joy.AtNeutralXY, JoystickPull := joy.AxisCmdY.DirectionPositive, JoystickPush := joy.AxisCmdY.DirectionNegative, BtnValidation := bench.Operator.JoyBtnRaw);
IF bench.Operator.JoyBtnRaw AND NOT previousButton THEN buttonEdges := buttonEdges + 1; END_IF; previousButton := bench.Operator.JoyBtnRaw;
ADVANCE_TIME(10000000);
bench(RawPosM1 := raw1, RawPosM2 := raw2);
joy(RawX := bench.Operator.JoyXRaw_ANA1, RawY := bench.Operator.JoyYRaw_ANA2, RawButton := bench.Operator.JoyBtnRaw, Cfg := cfg, NeutralXMem := nx, NeutralYMem := ny);
home(DeadmanArmed := joy.DeadmanArmed, JoystickDeflected := NOT joy.AtNeutralXY, JoystickPull := joy.AxisCmdY.DirectionPositive, JoystickPush := joy.AxisCmdY.DirectionNegative, BtnValidation := bench.Operator.JoyBtnRaw);
IF bench.Operator.JoyBtnRaw AND NOT previousButton THEN buttonEdges := buttonEdges + 1; END_IF; previousButton := bench.Operator.JoyBtnRaw;
ADVANCE_TIME(10000000);
bench(RawPosM1 := raw1, RawPosM2 := raw2);
joy(RawX := bench.Operator.JoyXRaw_ANA1, RawY := bench.Operator.JoyYRaw_ANA2, RawButton := bench.Operator.JoyBtnRaw, Cfg := cfg, NeutralXMem := nx, NeutralYMem := ny);
home(DeadmanArmed := joy.DeadmanArmed, JoystickDeflected := NOT joy.AtNeutralXY, JoystickPull := joy.AxisCmdY.DirectionPositive, JoystickPush := joy.AxisCmdY.DirectionNegative, BtnValidation := bench.Operator.JoyBtnRaw);
IF bench.Operator.JoyBtnRaw AND NOT previousButton THEN buttonEdges := buttonEdges + 1; END_IF; previousButton := bench.Operator.JoyBtnRaw;
ADVANCE_TIME(10000000);
bench(RawPosM1 := raw1, RawPosM2 := raw2);
joy(RawX := bench.Operator.JoyXRaw_ANA1, RawY := bench.Operator.JoyYRaw_ANA2, RawButton := bench.Operator.JoyBtnRaw, Cfg := cfg, NeutralXMem := nx, NeutralYMem := ny);
home(DeadmanArmed := joy.DeadmanArmed, JoystickDeflected := NOT joy.AtNeutralXY, JoystickPull := joy.AxisCmdY.DirectionPositive, JoystickPush := joy.AxisCmdY.DirectionNegative, BtnValidation := bench.Operator.JoyBtnRaw);
IF bench.Operator.JoyBtnRaw AND NOT previousButton THEN buttonEdges := buttonEdges + 1; END_IF; previousButton := bench.Operator.JoyBtnRaw;
ADVANCE_TIME(10000000);
bench(RawPosM1 := raw1, RawPosM2 := raw2);
joy(RawX := bench.Operator.JoyXRaw_ANA1, RawY := bench.Operator.JoyYRaw_ANA2, RawButton := bench.Operator.JoyBtnRaw, Cfg := cfg, NeutralXMem := nx, NeutralYMem := ny);
home(DeadmanArmed := joy.DeadmanArmed, JoystickDeflected := NOT joy.AtNeutralXY, JoystickPull := joy.AxisCmdY.DirectionPositive, JoystickPush := joy.AxisCmdY.DirectionNegative, BtnValidation := bench.Operator.JoyBtnRaw);
IF bench.Operator.JoyBtnRaw AND NOT previousButton THEN buttonEdges := buttonEdges + 1; END_IF; previousButton := bench.Operator.JoyBtnRaw;
ADVANCE_TIME(10000000);
bench(RawPosM1 := raw1, RawPosM2 := raw2);
joy(RawX := bench.Operator.JoyXRaw_ANA1, RawY := bench.Operator.JoyYRaw_ANA2, RawButton := bench.Operator.JoyBtnRaw, Cfg := cfg, NeutralXMem := nx, NeutralYMem := ny);
home(DeadmanArmed := joy.DeadmanArmed, JoystickDeflected := NOT joy.AtNeutralXY, JoystickPull := joy.AxisCmdY.DirectionPositive, JoystickPush := joy.AxisCmdY.DirectionNegative, BtnValidation := bench.Operator.JoyBtnRaw);
IF bench.Operator.JoyBtnRaw AND NOT previousButton THEN buttonEdges := buttonEdges + 1; END_IF; previousButton := bench.Operator.JoyBtnRaw;
ADVANCE_TIME(10000000);
bench(RawPosM1 := raw1, RawPosM2 := raw2);
joy(RawX := bench.Operator.JoyXRaw_ANA1, RawY := bench.Operator.JoyYRaw_ANA2, RawButton := bench.Operator.JoyBtnRaw, Cfg := cfg, NeutralXMem := nx, NeutralYMem := ny);
home(DeadmanArmed := joy.DeadmanArmed, JoystickDeflected := NOT joy.AtNeutralXY, JoystickPull := joy.AxisCmdY.DirectionPositive, JoystickPush := joy.AxisCmdY.DirectionNegative, BtnValidation := bench.Operator.JoyBtnRaw);
IF bench.Operator.JoyBtnRaw AND NOT previousButton THEN buttonEdges := buttonEdges + 1; END_IF; previousButton := bench.Operator.JoyBtnRaw;
ADVANCE_TIME(10000000);
bench(RawPosM1 := raw1, RawPosM2 := raw2);
joy(RawX := bench.Operator.JoyXRaw_ANA1, RawY := bench.Operator.JoyYRaw_ANA2, RawButton := bench.Operator.JoyBtnRaw, Cfg := cfg, NeutralXMem := nx, NeutralYMem := ny);
home(DeadmanArmed := joy.DeadmanArmed, JoystickDeflected := NOT joy.AtNeutralXY, JoystickPull := joy.AxisCmdY.DirectionPositive, JoystickPush := joy.AxisCmdY.DirectionNegative, BtnValidation := bench.Operator.JoyBtnRaw);
IF bench.Operator.JoyBtnRaw AND NOT previousButton THEN buttonEdges := buttonEdges + 1; END_IF; previousButton := bench.Operator.JoyBtnRaw;
ADVANCE_TIME(10000000);
bench(RawPosM1 := raw1, RawPosM2 := raw2);
joy(RawX := bench.Operator.JoyXRaw_ANA1, RawY := bench.Operator.JoyYRaw_ANA2, RawButton := bench.Operator.JoyBtnRaw, Cfg := cfg, NeutralXMem := nx, NeutralYMem := ny);
home(DeadmanArmed := joy.DeadmanArmed, JoystickDeflected := NOT joy.AtNeutralXY, JoystickPull := joy.AxisCmdY.DirectionPositive, JoystickPush := joy.AxisCmdY.DirectionNegative, BtnValidation := bench.Operator.JoyBtnRaw);
IF bench.Operator.JoyBtnRaw AND NOT previousButton THEN buttonEdges := buttonEdges + 1; END_IF; previousButton := bench.Operator.JoyBtnRaw;
ADVANCE_TIME(10000000);
bench(RawPosM1 := raw1, RawPosM2 := raw2);
joy(RawX := bench.Operator.JoyXRaw_ANA1, RawY := bench.Operator.JoyYRaw_ANA2, RawButton := bench.Operator.JoyBtnRaw, Cfg := cfg, NeutralXMem := nx, NeutralYMem := ny);
home(DeadmanArmed := joy.DeadmanArmed, JoystickDeflected := NOT joy.AtNeutralXY, JoystickPull := joy.AxisCmdY.DirectionPositive, JoystickPush := joy.AxisCmdY.DirectionNegative, BtnValidation := bench.Operator.JoyBtnRaw);
IF bench.Operator.JoyBtnRaw AND NOT previousButton THEN buttonEdges := buttonEdges + 1; END_IF; previousButton := bench.Operator.JoyBtnRaw;
ADVANCE_TIME(10000000);
bench(RawPosM1 := raw1, RawPosM2 := raw2);
joy(RawX := bench.Operator.JoyXRaw_ANA1, RawY := bench.Operator.JoyYRaw_ANA2, RawButton := bench.Operator.JoyBtnRaw, Cfg := cfg, NeutralXMem := nx, NeutralYMem := ny);
home(DeadmanArmed := joy.DeadmanArmed, JoystickDeflected := NOT joy.AtNeutralXY, JoystickPull := joy.AxisCmdY.DirectionPositive, JoystickPush := joy.AxisCmdY.DirectionNegative, BtnValidation := bench.Operator.JoyBtnRaw);
IF bench.Operator.JoyBtnRaw AND NOT previousButton THEN buttonEdges := buttonEdges + 1; END_IF; previousButton := bench.Operator.JoyBtnRaw;
ADVANCE_TIME(10000000);
bench(RawPosM1 := raw1, RawPosM2 := raw2);
joy(RawX := bench.Operator.JoyXRaw_ANA1, RawY := bench.Operator.JoyYRaw_ANA2, RawButton := bench.Operator.JoyBtnRaw, Cfg := cfg, NeutralXMem := nx, NeutralYMem := ny);
home(DeadmanArmed := joy.DeadmanArmed, JoystickDeflected := NOT joy.AtNeutralXY, JoystickPull := joy.AxisCmdY.DirectionPositive, JoystickPush := joy.AxisCmdY.DirectionNegative, BtnValidation := bench.Operator.JoyBtnRaw);
IF bench.Operator.JoyBtnRaw AND NOT previousButton THEN buttonEdges := buttonEdges + 1; END_IF; previousButton := bench.Operator.JoyBtnRaw;
ADVANCE_TIME(10000000);
bench(RawPosM1 := raw1, RawPosM2 := raw2);
joy(RawX := bench.Operator.JoyXRaw_ANA1, RawY := bench.Operator.JoyYRaw_ANA2, RawButton := bench.Operator.JoyBtnRaw, Cfg := cfg, NeutralXMem := nx, NeutralYMem := ny);
home(DeadmanArmed := joy.DeadmanArmed, JoystickDeflected := NOT joy.AtNeutralXY, JoystickPull := joy.AxisCmdY.DirectionPositive, JoystickPush := joy.AxisCmdY.DirectionNegative, BtnValidation := bench.Operator.JoyBtnRaw);
IF bench.Operator.JoyBtnRaw AND NOT previousButton THEN buttonEdges := buttonEdges + 1; END_IF; previousButton := bench.Operator.JoyBtnRaw;
ADVANCE_TIME(10000000);
bench(RawPosM1 := raw1, RawPosM2 := raw2);
joy(RawX := bench.Operator.JoyXRaw_ANA1, RawY := bench.Operator.JoyYRaw_ANA2, RawButton := bench.Operator.JoyBtnRaw, Cfg := cfg, NeutralXMem := nx, NeutralYMem := ny);
home(DeadmanArmed := joy.DeadmanArmed, JoystickDeflected := NOT joy.AtNeutralXY, JoystickPull := joy.AxisCmdY.DirectionPositive, JoystickPush := joy.AxisCmdY.DirectionNegative, BtnValidation := bench.Operator.JoyBtnRaw);
IF bench.Operator.JoyBtnRaw AND NOT previousButton THEN buttonEdges := buttonEdges + 1; END_IF; previousButton := bench.Operator.JoyBtnRaw;
ADVANCE_TIME(10000000);
bench(RawPosM1 := raw1, RawPosM2 := raw2);
joy(RawX := bench.Operator.JoyXRaw_ANA1, RawY := bench.Operator.JoyYRaw_ANA2, RawButton := bench.Operator.JoyBtnRaw, Cfg := cfg, NeutralXMem := nx, NeutralYMem := ny);
home(DeadmanArmed := joy.DeadmanArmed, JoystickDeflected := NOT joy.AtNeutralXY, JoystickPull := joy.AxisCmdY.DirectionPositive, JoystickPush := joy.AxisCmdY.DirectionNegative, BtnValidation := bench.Operator.JoyBtnRaw);
IF bench.Operator.JoyBtnRaw AND NOT previousButton THEN buttonEdges := buttonEdges + 1; END_IF; previousButton := bench.Operator.JoyBtnRaw;
ADVANCE_TIME(10000000);
bench(RawPosM1 := raw1, RawPosM2 := raw2);
joy(RawX := bench.Operator.JoyXRaw_ANA1, RawY := bench.Operator.JoyYRaw_ANA2, RawButton := bench.Operator.JoyBtnRaw, Cfg := cfg, NeutralXMem := nx, NeutralYMem := ny);
home(DeadmanArmed := joy.DeadmanArmed, JoystickDeflected := NOT joy.AtNeutralXY, JoystickPull := joy.AxisCmdY.DirectionPositive, JoystickPush := joy.AxisCmdY.DirectionNegative, BtnValidation := bench.Operator.JoyBtnRaw);
IF bench.Operator.JoyBtnRaw AND NOT previousButton THEN buttonEdges := buttonEdges + 1; END_IF; previousButton := bench.Operator.JoyBtnRaw;
ADVANCE_TIME(10000000);
bench(RawPosM1 := raw1, RawPosM2 := raw2);
joy(RawX := bench.Operator.JoyXRaw_ANA1, RawY := bench.Operator.JoyYRaw_ANA2, RawButton := bench.Operator.JoyBtnRaw, Cfg := cfg, NeutralXMem := nx, NeutralYMem := ny);
home(DeadmanArmed := joy.DeadmanArmed, JoystickDeflected := NOT joy.AtNeutralXY, JoystickPull := joy.AxisCmdY.DirectionPositive, JoystickPush := joy.AxisCmdY.DirectionNegative, BtnValidation := bench.Operator.JoyBtnRaw);
IF bench.Operator.JoyBtnRaw AND NOT previousButton THEN buttonEdges := buttonEdges + 1; END_IF; previousButton := bench.Operator.JoyBtnRaw;
ADVANCE_TIME(10000000);
bench(RawPosM1 := raw1, RawPosM2 := raw2);
joy(RawX := bench.Operator.JoyXRaw_ANA1, RawY := bench.Operator.JoyYRaw_ANA2, RawButton := bench.Operator.JoyBtnRaw, Cfg := cfg, NeutralXMem := nx, NeutralYMem := ny);
home(DeadmanArmed := joy.DeadmanArmed, JoystickDeflected := NOT joy.AtNeutralXY, JoystickPull := joy.AxisCmdY.DirectionPositive, JoystickPush := joy.AxisCmdY.DirectionNegative, BtnValidation := bench.Operator.JoyBtnRaw);
IF bench.Operator.JoyBtnRaw AND NOT previousButton THEN buttonEdges := buttonEdges + 1; END_IF; previousButton := bench.Operator.JoyBtnRaw;
ADVANCE_TIME(10000000);
bench(RawPosM1 := raw1, RawPosM2 := raw2);
joy(RawX := bench.Operator.JoyXRaw_ANA1, RawY := bench.Operator.JoyYRaw_ANA2, RawButton := bench.Operator.JoyBtnRaw, Cfg := cfg, NeutralXMem := nx, NeutralYMem := ny);
home(DeadmanArmed := joy.DeadmanArmed, JoystickDeflected := NOT joy.AtNeutralXY, JoystickPull := joy.AxisCmdY.DirectionPositive, JoystickPush := joy.AxisCmdY.DirectionNegative, BtnValidation := bench.Operator.JoyBtnRaw);
IF bench.Operator.JoyBtnRaw AND NOT previousButton THEN buttonEdges := buttonEdges + 1; END_IF; previousButton := bench.Operator.JoyBtnRaw;
ADVANCE_TIME(10000000);
bench(RawPosM1 := raw1, RawPosM2 := raw2);
joy(RawX := bench.Operator.JoyXRaw_ANA1, RawY := bench.Operator.JoyYRaw_ANA2, RawButton := bench.Operator.JoyBtnRaw, Cfg := cfg, NeutralXMem := nx, NeutralYMem := ny);
home(DeadmanArmed := joy.DeadmanArmed, JoystickDeflected := NOT joy.AtNeutralXY, JoystickPull := joy.AxisCmdY.DirectionPositive, JoystickPush := joy.AxisCmdY.DirectionNegative, BtnValidation := bench.Operator.JoyBtnRaw);
IF bench.Operator.JoyBtnRaw AND NOT previousButton THEN buttonEdges := buttonEdges + 1; END_IF; previousButton := bench.Operator.JoyBtnRaw;
ADVANCE_TIME(10000000);
bench(RawPosM1 := raw1, RawPosM2 := raw2);
joy(RawX := bench.Operator.JoyXRaw_ANA1, RawY := bench.Operator.JoyYRaw_ANA2, RawButton := bench.Operator.JoyBtnRaw, Cfg := cfg, NeutralXMem := nx, NeutralYMem := ny);
home(DeadmanArmed := joy.DeadmanArmed, JoystickDeflected := NOT joy.AtNeutralXY, JoystickPull := joy.AxisCmdY.DirectionPositive, JoystickPush := joy.AxisCmdY.DirectionNegative, BtnValidation := bench.Operator.JoyBtnRaw);
IF bench.Operator.JoyBtnRaw AND NOT previousButton THEN buttonEdges := buttonEdges + 1; END_IF; previousButton := bench.Operator.JoyBtnRaw;
ADVANCE_TIME(10000000);
bench(RawPosM1 := raw1, RawPosM2 := raw2);
joy(RawX := bench.Operator.JoyXRaw_ANA1, RawY := bench.Operator.JoyYRaw_ANA2, RawButton := bench.Operator.JoyBtnRaw, Cfg := cfg, NeutralXMem := nx, NeutralYMem := ny);
home(DeadmanArmed := joy.DeadmanArmed, JoystickDeflected := NOT joy.AtNeutralXY, JoystickPull := joy.AxisCmdY.DirectionPositive, JoystickPush := joy.AxisCmdY.DirectionNegative, BtnValidation := bench.Operator.JoyBtnRaw);
IF bench.Operator.JoyBtnRaw AND NOT previousButton THEN buttonEdges := buttonEdges + 1; END_IF; previousButton := bench.Operator.JoyBtnRaw;
ADVANCE_TIME(10000000);
bench(RawPosM1 := raw1, RawPosM2 := raw2);
joy(RawX := bench.Operator.JoyXRaw_ANA1, RawY := bench.Operator.JoyYRaw_ANA2, RawButton := bench.Operator.JoyBtnRaw, Cfg := cfg, NeutralXMem := nx, NeutralYMem := ny);
home(DeadmanArmed := joy.DeadmanArmed, JoystickDeflected := NOT joy.AtNeutralXY, JoystickPull := joy.AxisCmdY.DirectionPositive, JoystickPush := joy.AxisCmdY.DirectionNegative, BtnValidation := bench.Operator.JoyBtnRaw);
IF bench.Operator.JoyBtnRaw AND NOT previousButton THEN buttonEdges := buttonEdges + 1; END_IF; previousButton := bench.Operator.JoyBtnRaw;
ADVANCE_TIME(10000000);
bench(RawPosM1 := raw1, RawPosM2 := raw2);
joy(RawX := bench.Operator.JoyXRaw_ANA1, RawY := bench.Operator.JoyYRaw_ANA2, RawButton := bench.Operator.JoyBtnRaw, Cfg := cfg, NeutralXMem := nx, NeutralYMem := ny);
home(DeadmanArmed := joy.DeadmanArmed, JoystickDeflected := NOT joy.AtNeutralXY, JoystickPull := joy.AxisCmdY.DirectionPositive, JoystickPush := joy.AxisCmdY.DirectionNegative, BtnValidation := bench.Operator.JoyBtnRaw);
IF bench.Operator.JoyBtnRaw AND NOT previousButton THEN buttonEdges := buttonEdges + 1; END_IF; previousButton := bench.Operator.JoyBtnRaw;
ADVANCE_TIME(10000000);
bench(RawPosM1 := raw1, RawPosM2 := raw2);
joy(RawX := bench.Operator.JoyXRaw_ANA1, RawY := bench.Operator.JoyYRaw_ANA2, RawButton := bench.Operator.JoyBtnRaw, Cfg := cfg, NeutralXMem := nx, NeutralYMem := ny);
home(DeadmanArmed := joy.DeadmanArmed, JoystickDeflected := NOT joy.AtNeutralXY, JoystickPull := joy.AxisCmdY.DirectionPositive, JoystickPush := joy.AxisCmdY.DirectionNegative, BtnValidation := bench.Operator.JoyBtnRaw);
IF bench.Operator.JoyBtnRaw AND NOT previousButton THEN buttonEdges := buttonEdges + 1; END_IF; previousButton := bench.Operator.JoyBtnRaw;
ADVANCE_TIME(10000000);
bench(RawPosM1 := raw1, RawPosM2 := raw2);
joy(RawX := bench.Operator.JoyXRaw_ANA1, RawY := bench.Operator.JoyYRaw_ANA2, RawButton := bench.Operator.JoyBtnRaw, Cfg := cfg, NeutralXMem := nx, NeutralYMem := ny);
home(DeadmanArmed := joy.DeadmanArmed, JoystickDeflected := NOT joy.AtNeutralXY, JoystickPull := joy.AxisCmdY.DirectionPositive, JoystickPush := joy.AxisCmdY.DirectionNegative, BtnValidation := bench.Operator.JoyBtnRaw);
IF bench.Operator.JoyBtnRaw AND NOT previousButton THEN buttonEdges := buttonEdges + 1; END_IF; previousButton := bench.Operator.JoyBtnRaw;
ADVANCE_TIME(10000000);
bench(RawPosM1 := raw1, RawPosM2 := raw2);
joy(RawX := bench.Operator.JoyXRaw_ANA1, RawY := bench.Operator.JoyYRaw_ANA2, RawButton := bench.Operator.JoyBtnRaw, Cfg := cfg, NeutralXMem := nx, NeutralYMem := ny);
home(DeadmanArmed := joy.DeadmanArmed, JoystickDeflected := NOT joy.AtNeutralXY, JoystickPull := joy.AxisCmdY.DirectionPositive, JoystickPush := joy.AxisCmdY.DirectionNegative, BtnValidation := bench.Operator.JoyBtnRaw);
IF bench.Operator.JoyBtnRaw AND NOT previousButton THEN buttonEdges := buttonEdges + 1; END_IF; previousButton := bench.Operator.JoyBtnRaw;
ADVANCE_TIME(10000000);
bench(RawPosM1 := raw1, RawPosM2 := raw2);
joy(RawX := bench.Operator.JoyXRaw_ANA1, RawY := bench.Operator.JoyYRaw_ANA2, RawButton := bench.Operator.JoyBtnRaw, Cfg := cfg, NeutralXMem := nx, NeutralYMem := ny);
home(DeadmanArmed := joy.DeadmanArmed, JoystickDeflected := NOT joy.AtNeutralXY, JoystickPull := joy.AxisCmdY.DirectionPositive, JoystickPush := joy.AxisCmdY.DirectionNegative, BtnValidation := bench.Operator.JoyBtnRaw);
IF bench.Operator.JoyBtnRaw AND NOT previousButton THEN buttonEdges := buttonEdges + 1; END_IF; previousButton := bench.Operator.JoyBtnRaw;
ADVANCE_TIME(10000000);
bench(RawPosM1 := raw1, RawPosM2 := raw2);
joy(RawX := bench.Operator.JoyXRaw_ANA1, RawY := bench.Operator.JoyYRaw_ANA2, RawButton := bench.Operator.JoyBtnRaw, Cfg := cfg, NeutralXMem := nx, NeutralYMem := ny);
home(DeadmanArmed := joy.DeadmanArmed, JoystickDeflected := NOT joy.AtNeutralXY, JoystickPull := joy.AxisCmdY.DirectionPositive, JoystickPush := joy.AxisCmdY.DirectionNegative, BtnValidation := bench.Operator.JoyBtnRaw);
IF bench.Operator.JoyBtnRaw AND NOT previousButton THEN buttonEdges := buttonEdges + 1; END_IF; previousButton := bench.Operator.JoyBtnRaw;
ADVANCE_TIME(10000000);
bench(RawPosM1 := raw1, RawPosM2 := raw2);
joy(RawX := bench.Operator.JoyXRaw_ANA1, RawY := bench.Operator.JoyYRaw_ANA2, RawButton := bench.Operator.JoyBtnRaw, Cfg := cfg, NeutralXMem := nx, NeutralYMem := ny);
home(DeadmanArmed := joy.DeadmanArmed, JoystickDeflected := NOT joy.AtNeutralXY, JoystickPull := joy.AxisCmdY.DirectionPositive, JoystickPush := joy.AxisCmdY.DirectionNegative, BtnValidation := bench.Operator.JoyBtnRaw);
IF bench.Operator.JoyBtnRaw AND NOT previousButton THEN buttonEdges := buttonEdges + 1; END_IF; previousButton := bench.Operator.JoyBtnRaw;
ADVANCE_TIME(10000000);
bench(RawPosM1 := raw1, RawPosM2 := raw2);
joy(RawX := bench.Operator.JoyXRaw_ANA1, RawY := bench.Operator.JoyYRaw_ANA2, RawButton := bench.Operator.JoyBtnRaw, Cfg := cfg, NeutralXMem := nx, NeutralYMem := ny);
home(DeadmanArmed := joy.DeadmanArmed, JoystickDeflected := NOT joy.AtNeutralXY, JoystickPull := joy.AxisCmdY.DirectionPositive, JoystickPush := joy.AxisCmdY.DirectionNegative, BtnValidation := bench.Operator.JoyBtnRaw);
IF bench.Operator.JoyBtnRaw AND NOT previousButton THEN buttonEdges := buttonEdges + 1; END_IF; previousButton := bench.Operator.JoyBtnRaw;
ADVANCE_TIME(10000000);
bench(RawPosM1 := raw1, RawPosM2 := raw2);
joy(RawX := bench.Operator.JoyXRaw_ANA1, RawY := bench.Operator.JoyYRaw_ANA2, RawButton := bench.Operator.JoyBtnRaw, Cfg := cfg, NeutralXMem := nx, NeutralYMem := ny);
home(DeadmanArmed := joy.DeadmanArmed, JoystickDeflected := NOT joy.AtNeutralXY, JoystickPull := joy.AxisCmdY.DirectionPositive, JoystickPush := joy.AxisCmdY.DirectionNegative, BtnValidation := bench.Operator.JoyBtnRaw);
IF bench.Operator.JoyBtnRaw AND NOT previousButton THEN buttonEdges := buttonEdges + 1; END_IF; previousButton := bench.Operator.JoyBtnRaw;
ADVANCE_TIME(10000000);
bench(RawPosM1 := raw1, RawPosM2 := raw2);
joy(RawX := bench.Operator.JoyXRaw_ANA1, RawY := bench.Operator.JoyYRaw_ANA2, RawButton := bench.Operator.JoyBtnRaw, Cfg := cfg, NeutralXMem := nx, NeutralYMem := ny);
home(DeadmanArmed := joy.DeadmanArmed, JoystickDeflected := NOT joy.AtNeutralXY, JoystickPull := joy.AxisCmdY.DirectionPositive, JoystickPush := joy.AxisCmdY.DirectionNegative, BtnValidation := bench.Operator.JoyBtnRaw);
IF bench.Operator.JoyBtnRaw AND NOT previousButton THEN buttonEdges := buttonEdges + 1; END_IF; previousButton := bench.Operator.JoyBtnRaw;
ASSERT_TRUE(joy.AxisCmdY.StartStop, 'Geste initial effectif');
joy.ArmingPermit := FALSE;
ADVANCE_TIME(10000000);
bench(RawPosM1 := raw1, RawPosM2 := raw2);
joy(RawX := bench.Operator.JoyXRaw_ANA1, RawY := bench.Operator.JoyYRaw_ANA2, RawButton := bench.Operator.JoyBtnRaw, Cfg := cfg, NeutralXMem := nx, NeutralYMem := ny);
home(DeadmanArmed := joy.DeadmanArmed, JoystickDeflected := NOT joy.AtNeutralXY, JoystickPull := joy.AxisCmdY.DirectionPositive, JoystickPush := joy.AxisCmdY.DirectionNegative, BtnValidation := bench.Operator.JoyBtnRaw);
IF bench.Operator.JoyBtnRaw AND NOT previousButton THEN buttonEdges := buttonEdges + 1; END_IF; previousButton := bench.Operator.JoyBtnRaw;
ASSERT_FALSE(joy.DeadmanArmed, 'Desarmement immediat reel');
joy.ArmingPermit := TRUE;
ADVANCE_TIME(10000000);
bench(RawPosM1 := raw1, RawPosM2 := raw2);
joy(RawX := bench.Operator.JoyXRaw_ANA1, RawY := bench.Operator.JoyYRaw_ANA2, RawButton := bench.Operator.JoyBtnRaw, Cfg := cfg, NeutralXMem := nx, NeutralYMem := ny);
home(DeadmanArmed := joy.DeadmanArmed, JoystickDeflected := NOT joy.AtNeutralXY, JoystickPull := joy.AxisCmdY.DirectionPositive, JoystickPush := joy.AxisCmdY.DirectionNegative, BtnValidation := bench.Operator.JoyBtnRaw);
IF bench.Operator.JoyBtnRaw AND NOT previousButton THEN buttonEdges := buttonEdges + 1; END_IF; previousButton := bench.Operator.JoyBtnRaw;
ASSERT_FALSE(joy.AxisCmdY.StartStop, 'Pas de reprise automatique');
ADVANCE_TIME(10000000);
bench(RawPosM1 := raw1, RawPosM2 := raw2);
joy(RawX := bench.Operator.JoyXRaw_ANA1, RawY := bench.Operator.JoyYRaw_ANA2, RawButton := bench.Operator.JoyBtnRaw, Cfg := cfg, NeutralXMem := nx, NeutralYMem := ny);
home(DeadmanArmed := joy.DeadmanArmed, JoystickDeflected := NOT joy.AtNeutralXY, JoystickPull := joy.AxisCmdY.DirectionPositive, JoystickPush := joy.AxisCmdY.DirectionNegative, BtnValidation := bench.Operator.JoyBtnRaw);
IF bench.Operator.JoyBtnRaw AND NOT previousButton THEN buttonEdges := buttonEdges + 1; END_IF; previousButton := bench.Operator.JoyBtnRaw;
ASSERT_FALSE(joy.AxisCmdY.StartStop, 'Pas de reprise automatique');
ADVANCE_TIME(10000000);
bench(RawPosM1 := raw1, RawPosM2 := raw2);
joy(RawX := bench.Operator.JoyXRaw_ANA1, RawY := bench.Operator.JoyYRaw_ANA2, RawButton := bench.Operator.JoyBtnRaw, Cfg := cfg, NeutralXMem := nx, NeutralYMem := ny);
home(DeadmanArmed := joy.DeadmanArmed, JoystickDeflected := NOT joy.AtNeutralXY, JoystickPull := joy.AxisCmdY.DirectionPositive, JoystickPush := joy.AxisCmdY.DirectionNegative, BtnValidation := bench.Operator.JoyBtnRaw);
IF bench.Operator.JoyBtnRaw AND NOT previousButton THEN buttonEdges := buttonEdges + 1; END_IF; previousButton := bench.Operator.JoyBtnRaw;
ASSERT_FALSE(joy.AxisCmdY.StartStop, 'Pas de reprise automatique');
ADVANCE_TIME(10000000);
bench(RawPosM1 := raw1, RawPosM2 := raw2);
joy(RawX := bench.Operator.JoyXRaw_ANA1, RawY := bench.Operator.JoyYRaw_ANA2, RawButton := bench.Operator.JoyBtnRaw, Cfg := cfg, NeutralXMem := nx, NeutralYMem := ny);
home(DeadmanArmed := joy.DeadmanArmed, JoystickDeflected := NOT joy.AtNeutralXY, JoystickPull := joy.AxisCmdY.DirectionPositive, JoystickPush := joy.AxisCmdY.DirectionNegative, BtnValidation := bench.Operator.JoyBtnRaw);
IF bench.Operator.JoyBtnRaw AND NOT previousButton THEN buttonEdges := buttonEdges + 1; END_IF; previousButton := bench.Operator.JoyBtnRaw;
ASSERT_FALSE(joy.AxisCmdY.StartStop, 'Pas de reprise automatique');
ADVANCE_TIME(10000000);
bench(RawPosM1 := raw1, RawPosM2 := raw2);
joy(RawX := bench.Operator.JoyXRaw_ANA1, RawY := bench.Operator.JoyYRaw_ANA2, RawButton := bench.Operator.JoyBtnRaw, Cfg := cfg, NeutralXMem := nx, NeutralYMem := ny);
home(DeadmanArmed := joy.DeadmanArmed, JoystickDeflected := NOT joy.AtNeutralXY, JoystickPull := joy.AxisCmdY.DirectionPositive, JoystickPush := joy.AxisCmdY.DirectionNegative, BtnValidation := bench.Operator.JoyBtnRaw);
IF bench.Operator.JoyBtnRaw AND NOT previousButton THEN buttonEdges := buttonEdges + 1; END_IF; previousButton := bench.Operator.JoyBtnRaw;
ASSERT_FALSE(joy.AxisCmdY.StartStop, 'Pas de reprise automatique');
ADVANCE_TIME(10000000);
bench(RawPosM1 := raw1, RawPosM2 := raw2);
joy(RawX := bench.Operator.JoyXRaw_ANA1, RawY := bench.Operator.JoyYRaw_ANA2, RawButton := bench.Operator.JoyBtnRaw, Cfg := cfg, NeutralXMem := nx, NeutralYMem := ny);
home(DeadmanArmed := joy.DeadmanArmed, JoystickDeflected := NOT joy.AtNeutralXY, JoystickPull := joy.AxisCmdY.DirectionPositive, JoystickPush := joy.AxisCmdY.DirectionNegative, BtnValidation := bench.Operator.JoyBtnRaw);
IF bench.Operator.JoyBtnRaw AND NOT previousButton THEN buttonEdges := buttonEdges + 1; END_IF; previousButton := bench.Operator.JoyBtnRaw;
ASSERT_FALSE(joy.AxisCmdY.StartStop, 'Pas de reprise automatique');
ADVANCE_TIME(10000000);
bench(RawPosM1 := raw1, RawPosM2 := raw2);
joy(RawX := bench.Operator.JoyXRaw_ANA1, RawY := bench.Operator.JoyYRaw_ANA2, RawButton := bench.Operator.JoyBtnRaw, Cfg := cfg, NeutralXMem := nx, NeutralYMem := ny);
home(DeadmanArmed := joy.DeadmanArmed, JoystickDeflected := NOT joy.AtNeutralXY, JoystickPull := joy.AxisCmdY.DirectionPositive, JoystickPush := joy.AxisCmdY.DirectionNegative, BtnValidation := bench.Operator.JoyBtnRaw);
IF bench.Operator.JoyBtnRaw AND NOT previousButton THEN buttonEdges := buttonEdges + 1; END_IF; previousButton := bench.Operator.JoyBtnRaw;
ASSERT_FALSE(joy.AxisCmdY.StartStop, 'Pas de reprise automatique');
ADVANCE_TIME(10000000);
bench(RawPosM1 := raw1, RawPosM2 := raw2);
joy(RawX := bench.Operator.JoyXRaw_ANA1, RawY := bench.Operator.JoyYRaw_ANA2, RawButton := bench.Operator.JoyBtnRaw, Cfg := cfg, NeutralXMem := nx, NeutralYMem := ny);
home(DeadmanArmed := joy.DeadmanArmed, JoystickDeflected := NOT joy.AtNeutralXY, JoystickPull := joy.AxisCmdY.DirectionPositive, JoystickPush := joy.AxisCmdY.DirectionNegative, BtnValidation := bench.Operator.JoyBtnRaw);
IF bench.Operator.JoyBtnRaw AND NOT previousButton THEN buttonEdges := buttonEdges + 1; END_IF; previousButton := bench.Operator.JoyBtnRaw;
ASSERT_FALSE(joy.AxisCmdY.StartStop, 'Pas de reprise automatique');
ADVANCE_TIME(10000000);
bench(RawPosM1 := raw1, RawPosM2 := raw2);
joy(RawX := bench.Operator.JoyXRaw_ANA1, RawY := bench.Operator.JoyYRaw_ANA2, RawButton := bench.Operator.JoyBtnRaw, Cfg := cfg, NeutralXMem := nx, NeutralYMem := ny);
home(DeadmanArmed := joy.DeadmanArmed, JoystickDeflected := NOT joy.AtNeutralXY, JoystickPull := joy.AxisCmdY.DirectionPositive, JoystickPush := joy.AxisCmdY.DirectionNegative, BtnValidation := bench.Operator.JoyBtnRaw);
IF bench.Operator.JoyBtnRaw AND NOT previousButton THEN buttonEdges := buttonEdges + 1; END_IF; previousButton := bench.Operator.JoyBtnRaw;
ASSERT_FALSE(joy.AxisCmdY.StartStop, 'Pas de reprise automatique');
ADVANCE_TIME(10000000);
bench(RawPosM1 := raw1, RawPosM2 := raw2);
joy(RawX := bench.Operator.JoyXRaw_ANA1, RawY := bench.Operator.JoyYRaw_ANA2, RawButton := bench.Operator.JoyBtnRaw, Cfg := cfg, NeutralXMem := nx, NeutralYMem := ny);
home(DeadmanArmed := joy.DeadmanArmed, JoystickDeflected := NOT joy.AtNeutralXY, JoystickPull := joy.AxisCmdY.DirectionPositive, JoystickPush := joy.AxisCmdY.DirectionNegative, BtnValidation := bench.Operator.JoyBtnRaw);
IF bench.Operator.JoyBtnRaw AND NOT previousButton THEN buttonEdges := buttonEdges + 1; END_IF; previousButton := bench.Operator.JoyBtnRaw;
ASSERT_FALSE(joy.AxisCmdY.StartStop, 'Pas de reprise automatique');
ADVANCE_TIME(10000000);
bench(RawPosM1 := raw1, RawPosM2 := raw2);
joy(RawX := bench.Operator.JoyXRaw_ANA1, RawY := bench.Operator.JoyYRaw_ANA2, RawButton := bench.Operator.JoyBtnRaw, Cfg := cfg, NeutralXMem := nx, NeutralYMem := ny);
home(DeadmanArmed := joy.DeadmanArmed, JoystickDeflected := NOT joy.AtNeutralXY, JoystickPull := joy.AxisCmdY.DirectionPositive, JoystickPush := joy.AxisCmdY.DirectionNegative, BtnValidation := bench.Operator.JoyBtnRaw);
IF bench.Operator.JoyBtnRaw AND NOT previousButton THEN buttonEdges := buttonEdges + 1; END_IF; previousButton := bench.Operator.JoyBtnRaw;
ASSERT_FALSE(joy.AxisCmdY.StartStop, 'Pas de reprise automatique');
ADVANCE_TIME(10000000);
bench(RawPosM1 := raw1, RawPosM2 := raw2);
joy(RawX := bench.Operator.JoyXRaw_ANA1, RawY := bench.Operator.JoyYRaw_ANA2, RawButton := bench.Operator.JoyBtnRaw, Cfg := cfg, NeutralXMem := nx, NeutralYMem := ny);
home(DeadmanArmed := joy.DeadmanArmed, JoystickDeflected := NOT joy.AtNeutralXY, JoystickPull := joy.AxisCmdY.DirectionPositive, JoystickPush := joy.AxisCmdY.DirectionNegative, BtnValidation := bench.Operator.JoyBtnRaw);
IF bench.Operator.JoyBtnRaw AND NOT previousButton THEN buttonEdges := buttonEdges + 1; END_IF; previousButton := bench.Operator.JoyBtnRaw;
ASSERT_FALSE(joy.AxisCmdY.StartStop, 'Pas de reprise automatique');
ADVANCE_TIME(10000000);
bench(RawPosM1 := raw1, RawPosM2 := raw2);
joy(RawX := bench.Operator.JoyXRaw_ANA1, RawY := bench.Operator.JoyYRaw_ANA2, RawButton := bench.Operator.JoyBtnRaw, Cfg := cfg, NeutralXMem := nx, NeutralYMem := ny);
home(DeadmanArmed := joy.DeadmanArmed, JoystickDeflected := NOT joy.AtNeutralXY, JoystickPull := joy.AxisCmdY.DirectionPositive, JoystickPush := joy.AxisCmdY.DirectionNegative, BtnValidation := bench.Operator.JoyBtnRaw);
IF bench.Operator.JoyBtnRaw AND NOT previousButton THEN buttonEdges := buttonEdges + 1; END_IF; previousButton := bench.Operator.JoyBtnRaw;
ASSERT_FALSE(joy.AxisCmdY.StartStop, 'Pas de reprise automatique');
ADVANCE_TIME(10000000);
bench(RawPosM1 := raw1, RawPosM2 := raw2);
joy(RawX := bench.Operator.JoyXRaw_ANA1, RawY := bench.Operator.JoyYRaw_ANA2, RawButton := bench.Operator.JoyBtnRaw, Cfg := cfg, NeutralXMem := nx, NeutralYMem := ny);
home(DeadmanArmed := joy.DeadmanArmed, JoystickDeflected := NOT joy.AtNeutralXY, JoystickPull := joy.AxisCmdY.DirectionPositive, JoystickPush := joy.AxisCmdY.DirectionNegative, BtnValidation := bench.Operator.JoyBtnRaw);
IF bench.Operator.JoyBtnRaw AND NOT previousButton THEN buttonEdges := buttonEdges + 1; END_IF; previousButton := bench.Operator.JoyBtnRaw;
ASSERT_FALSE(joy.AxisCmdY.StartStop, 'Pas de reprise automatique');
ADVANCE_TIME(10000000);
bench(RawPosM1 := raw1, RawPosM2 := raw2);
joy(RawX := bench.Operator.JoyXRaw_ANA1, RawY := bench.Operator.JoyYRaw_ANA2, RawButton := bench.Operator.JoyBtnRaw, Cfg := cfg, NeutralXMem := nx, NeutralYMem := ny);
home(DeadmanArmed := joy.DeadmanArmed, JoystickDeflected := NOT joy.AtNeutralXY, JoystickPull := joy.AxisCmdY.DirectionPositive, JoystickPush := joy.AxisCmdY.DirectionNegative, BtnValidation := bench.Operator.JoyBtnRaw);
IF bench.Operator.JoyBtnRaw AND NOT previousButton THEN buttonEdges := buttonEdges + 1; END_IF; previousButton := bench.Operator.JoyBtnRaw;
ASSERT_FALSE(joy.AxisCmdY.StartStop, 'Pas de reprise automatique');
ADVANCE_TIME(10000000);
bench(RawPosM1 := raw1, RawPosM2 := raw2);
joy(RawX := bench.Operator.JoyXRaw_ANA1, RawY := bench.Operator.JoyYRaw_ANA2, RawButton := bench.Operator.JoyBtnRaw, Cfg := cfg, NeutralXMem := nx, NeutralYMem := ny);
home(DeadmanArmed := joy.DeadmanArmed, JoystickDeflected := NOT joy.AtNeutralXY, JoystickPull := joy.AxisCmdY.DirectionPositive, JoystickPush := joy.AxisCmdY.DirectionNegative, BtnValidation := bench.Operator.JoyBtnRaw);
IF bench.Operator.JoyBtnRaw AND NOT previousButton THEN buttonEdges := buttonEdges + 1; END_IF; previousButton := bench.Operator.JoyBtnRaw;
ASSERT_FALSE(joy.AxisCmdY.StartStop, 'Pas de reprise automatique');
ADVANCE_TIME(10000000);
bench(RawPosM1 := raw1, RawPosM2 := raw2);
joy(RawX := bench.Operator.JoyXRaw_ANA1, RawY := bench.Operator.JoyYRaw_ANA2, RawButton := bench.Operator.JoyBtnRaw, Cfg := cfg, NeutralXMem := nx, NeutralYMem := ny);
home(DeadmanArmed := joy.DeadmanArmed, JoystickDeflected := NOT joy.AtNeutralXY, JoystickPull := joy.AxisCmdY.DirectionPositive, JoystickPush := joy.AxisCmdY.DirectionNegative, BtnValidation := bench.Operator.JoyBtnRaw);
IF bench.Operator.JoyBtnRaw AND NOT previousButton THEN buttonEdges := buttonEdges + 1; END_IF; previousButton := bench.Operator.JoyBtnRaw;
ASSERT_FALSE(joy.AxisCmdY.StartStop, 'Pas de reprise automatique');
ADVANCE_TIME(10000000);
bench(RawPosM1 := raw1, RawPosM2 := raw2);
joy(RawX := bench.Operator.JoyXRaw_ANA1, RawY := bench.Operator.JoyYRaw_ANA2, RawButton := bench.Operator.JoyBtnRaw, Cfg := cfg, NeutralXMem := nx, NeutralYMem := ny);
home(DeadmanArmed := joy.DeadmanArmed, JoystickDeflected := NOT joy.AtNeutralXY, JoystickPull := joy.AxisCmdY.DirectionPositive, JoystickPush := joy.AxisCmdY.DirectionNegative, BtnValidation := bench.Operator.JoyBtnRaw);
IF bench.Operator.JoyBtnRaw AND NOT previousButton THEN buttonEdges := buttonEdges + 1; END_IF; previousButton := bench.Operator.JoyBtnRaw;
ASSERT_FALSE(joy.AxisCmdY.StartStop, 'Pas de reprise automatique');
ADVANCE_TIME(10000000);
bench(RawPosM1 := raw1, RawPosM2 := raw2);
joy(RawX := bench.Operator.JoyXRaw_ANA1, RawY := bench.Operator.JoyYRaw_ANA2, RawButton := bench.Operator.JoyBtnRaw, Cfg := cfg, NeutralXMem := nx, NeutralYMem := ny);
home(DeadmanArmed := joy.DeadmanArmed, JoystickDeflected := NOT joy.AtNeutralXY, JoystickPull := joy.AxisCmdY.DirectionPositive, JoystickPush := joy.AxisCmdY.DirectionNegative, BtnValidation := bench.Operator.JoyBtnRaw);
IF bench.Operator.JoyBtnRaw AND NOT previousButton THEN buttonEdges := buttonEdges + 1; END_IF; previousButton := bench.Operator.JoyBtnRaw;
ASSERT_FALSE(joy.AxisCmdY.StartStop, 'Pas de reprise automatique');
ADVANCE_TIME(10000000);
bench(RawPosM1 := raw1, RawPosM2 := raw2);
joy(RawX := bench.Operator.JoyXRaw_ANA1, RawY := bench.Operator.JoyYRaw_ANA2, RawButton := bench.Operator.JoyBtnRaw, Cfg := cfg, NeutralXMem := nx, NeutralYMem := ny);
home(DeadmanArmed := joy.DeadmanArmed, JoystickDeflected := NOT joy.AtNeutralXY, JoystickPull := joy.AxisCmdY.DirectionPositive, JoystickPush := joy.AxisCmdY.DirectionNegative, BtnValidation := bench.Operator.JoyBtnRaw);
IF bench.Operator.JoyBtnRaw AND NOT previousButton THEN buttonEdges := buttonEdges + 1; END_IF; previousButton := bench.Operator.JoyBtnRaw;
ASSERT_FALSE(joy.AxisCmdY.StartStop, 'Pas de reprise automatique');
ADVANCE_TIME(10000000);
bench(RawPosM1 := raw1, RawPosM2 := raw2);
joy(RawX := bench.Operator.JoyXRaw_ANA1, RawY := bench.Operator.JoyYRaw_ANA2, RawButton := bench.Operator.JoyBtnRaw, Cfg := cfg, NeutralXMem := nx, NeutralYMem := ny);
home(DeadmanArmed := joy.DeadmanArmed, JoystickDeflected := NOT joy.AtNeutralXY, JoystickPull := joy.AxisCmdY.DirectionPositive, JoystickPush := joy.AxisCmdY.DirectionNegative, BtnValidation := bench.Operator.JoyBtnRaw);
IF bench.Operator.JoyBtnRaw AND NOT previousButton THEN buttonEdges := buttonEdges + 1; END_IF; previousButton := bench.Operator.JoyBtnRaw;
ASSERT_FALSE(joy.AxisCmdY.StartStop, 'Pas de reprise automatique');
ADVANCE_TIME(10000000);
bench(RawPosM1 := raw1, RawPosM2 := raw2);
joy(RawX := bench.Operator.JoyXRaw_ANA1, RawY := bench.Operator.JoyYRaw_ANA2, RawButton := bench.Operator.JoyBtnRaw, Cfg := cfg, NeutralXMem := nx, NeutralYMem := ny);
home(DeadmanArmed := joy.DeadmanArmed, JoystickDeflected := NOT joy.AtNeutralXY, JoystickPull := joy.AxisCmdY.DirectionPositive, JoystickPush := joy.AxisCmdY.DirectionNegative, BtnValidation := bench.Operator.JoyBtnRaw);
IF bench.Operator.JoyBtnRaw AND NOT previousButton THEN buttonEdges := buttonEdges + 1; END_IF; previousButton := bench.Operator.JoyBtnRaw;
ASSERT_FALSE(joy.AxisCmdY.StartStop, 'Pas de reprise automatique');
ADVANCE_TIME(10000000);
bench(RawPosM1 := raw1, RawPosM2 := raw2);
joy(RawX := bench.Operator.JoyXRaw_ANA1, RawY := bench.Operator.JoyYRaw_ANA2, RawButton := bench.Operator.JoyBtnRaw, Cfg := cfg, NeutralXMem := nx, NeutralYMem := ny);
home(DeadmanArmed := joy.DeadmanArmed, JoystickDeflected := NOT joy.AtNeutralXY, JoystickPull := joy.AxisCmdY.DirectionPositive, JoystickPush := joy.AxisCmdY.DirectionNegative, BtnValidation := bench.Operator.JoyBtnRaw);
IF bench.Operator.JoyBtnRaw AND NOT previousButton THEN buttonEdges := buttonEdges + 1; END_IF; previousButton := bench.Operator.JoyBtnRaw;
ASSERT_FALSE(joy.AxisCmdY.StartStop, 'Pas de reprise automatique');
ADVANCE_TIME(10000000);
bench(RawPosM1 := raw1, RawPosM2 := raw2);
joy(RawX := bench.Operator.JoyXRaw_ANA1, RawY := bench.Operator.JoyYRaw_ANA2, RawButton := bench.Operator.JoyBtnRaw, Cfg := cfg, NeutralXMem := nx, NeutralYMem := ny);
home(DeadmanArmed := joy.DeadmanArmed, JoystickDeflected := NOT joy.AtNeutralXY, JoystickPull := joy.AxisCmdY.DirectionPositive, JoystickPush := joy.AxisCmdY.DirectionNegative, BtnValidation := bench.Operator.JoyBtnRaw);
IF bench.Operator.JoyBtnRaw AND NOT previousButton THEN buttonEdges := buttonEdges + 1; END_IF; previousButton := bench.Operator.JoyBtnRaw;
ASSERT_FALSE(joy.AxisCmdY.StartStop, 'Pas de reprise automatique');
ADVANCE_TIME(10000000);
bench(RawPosM1 := raw1, RawPosM2 := raw2);
joy(RawX := bench.Operator.JoyXRaw_ANA1, RawY := bench.Operator.JoyYRaw_ANA2, RawButton := bench.Operator.JoyBtnRaw, Cfg := cfg, NeutralXMem := nx, NeutralYMem := ny);
home(DeadmanArmed := joy.DeadmanArmed, JoystickDeflected := NOT joy.AtNeutralXY, JoystickPull := joy.AxisCmdY.DirectionPositive, JoystickPush := joy.AxisCmdY.DirectionNegative, BtnValidation := bench.Operator.JoyBtnRaw);
IF bench.Operator.JoyBtnRaw AND NOT previousButton THEN buttonEdges := buttonEdges + 1; END_IF; previousButton := bench.Operator.JoyBtnRaw;
ASSERT_FALSE(joy.AxisCmdY.StartStop, 'Pas de reprise automatique');
ADVANCE_TIME(10000000);
bench(RawPosM1 := raw1, RawPosM2 := raw2);
joy(RawX := bench.Operator.JoyXRaw_ANA1, RawY := bench.Operator.JoyYRaw_ANA2, RawButton := bench.Operator.JoyBtnRaw, Cfg := cfg, NeutralXMem := nx, NeutralYMem := ny);
home(DeadmanArmed := joy.DeadmanArmed, JoystickDeflected := NOT joy.AtNeutralXY, JoystickPull := joy.AxisCmdY.DirectionPositive, JoystickPush := joy.AxisCmdY.DirectionNegative, BtnValidation := bench.Operator.JoyBtnRaw);
IF bench.Operator.JoyBtnRaw AND NOT previousButton THEN buttonEdges := buttonEdges + 1; END_IF; previousButton := bench.Operator.JoyBtnRaw;
ASSERT_FALSE(joy.AxisCmdY.StartStop, 'Pas de reprise automatique');
ADVANCE_TIME(10000000);
bench(RawPosM1 := raw1, RawPosM2 := raw2);
joy(RawX := bench.Operator.JoyXRaw_ANA1, RawY := bench.Operator.JoyYRaw_ANA2, RawButton := bench.Operator.JoyBtnRaw, Cfg := cfg, NeutralXMem := nx, NeutralYMem := ny);
home(DeadmanArmed := joy.DeadmanArmed, JoystickDeflected := NOT joy.AtNeutralXY, JoystickPull := joy.AxisCmdY.DirectionPositive, JoystickPush := joy.AxisCmdY.DirectionNegative, BtnValidation := bench.Operator.JoyBtnRaw);
IF bench.Operator.JoyBtnRaw AND NOT previousButton THEN buttonEdges := buttonEdges + 1; END_IF; previousButton := bench.Operator.JoyBtnRaw;
ASSERT_FALSE(joy.AxisCmdY.StartStop, 'Pas de reprise automatique');
ADVANCE_TIME(10000000);
bench(RawPosM1 := raw1, RawPosM2 := raw2);
joy(RawX := bench.Operator.JoyXRaw_ANA1, RawY := bench.Operator.JoyYRaw_ANA2, RawButton := bench.Operator.JoyBtnRaw, Cfg := cfg, NeutralXMem := nx, NeutralYMem := ny);
home(DeadmanArmed := joy.DeadmanArmed, JoystickDeflected := NOT joy.AtNeutralXY, JoystickPull := joy.AxisCmdY.DirectionPositive, JoystickPush := joy.AxisCmdY.DirectionNegative, BtnValidation := bench.Operator.JoyBtnRaw);
IF bench.Operator.JoyBtnRaw AND NOT previousButton THEN buttonEdges := buttonEdges + 1; END_IF; previousButton := bench.Operator.JoyBtnRaw;
ASSERT_FALSE(joy.AxisCmdY.StartStop, 'Pas de reprise automatique');
ADVANCE_TIME(10000000);
bench(RawPosM1 := raw1, RawPosM2 := raw2);
joy(RawX := bench.Operator.JoyXRaw_ANA1, RawY := bench.Operator.JoyYRaw_ANA2, RawButton := bench.Operator.JoyBtnRaw, Cfg := cfg, NeutralXMem := nx, NeutralYMem := ny);
home(DeadmanArmed := joy.DeadmanArmed, JoystickDeflected := NOT joy.AtNeutralXY, JoystickPull := joy.AxisCmdY.DirectionPositive, JoystickPush := joy.AxisCmdY.DirectionNegative, BtnValidation := bench.Operator.JoyBtnRaw);
IF bench.Operator.JoyBtnRaw AND NOT previousButton THEN buttonEdges := buttonEdges + 1; END_IF; previousButton := bench.Operator.JoyBtnRaw;
ASSERT_FALSE(joy.AxisCmdY.StartStop, 'Pas de reprise automatique');
ADVANCE_TIME(10000000);
bench(RawPosM1 := raw1, RawPosM2 := raw2);
joy(RawX := bench.Operator.JoyXRaw_ANA1, RawY := bench.Operator.JoyYRaw_ANA2, RawButton := bench.Operator.JoyBtnRaw, Cfg := cfg, NeutralXMem := nx, NeutralYMem := ny);
home(DeadmanArmed := joy.DeadmanArmed, JoystickDeflected := NOT joy.AtNeutralXY, JoystickPull := joy.AxisCmdY.DirectionPositive, JoystickPush := joy.AxisCmdY.DirectionNegative, BtnValidation := bench.Operator.JoyBtnRaw);
IF bench.Operator.JoyBtnRaw AND NOT previousButton THEN buttonEdges := buttonEdges + 1; END_IF; previousButton := bench.Operator.JoyBtnRaw;
ASSERT_FALSE(joy.AxisCmdY.StartStop, 'Pas de reprise automatique');
ASSERT_EQ(buttonEdges, 1, 'Pas de nouveau front simule');
END_TEST
